(* IEC 61131-3 sources: iecf/harness/cases (part 3) *)

(* ---- locmore.st ---- *)
(* Located variables without a name (Ed.3 Loc_Var_Decl: Variable_Name ?)
   and a FOR control variable at an address. Worked by hand:
   AT %QW4 : INT := 5 sets %QW4 to 5 (Q bytes 4, 5: 05 00) as the
   program is set up; AT %MB0 : ARRAY [1..2] OF BYTE := [1, 2] sets
   %MB0, %MB1 (01 02); AT %QB9 : BYTE := 7 sets %QB9 (07) -
   in the PROGRAM: a block's VAR has no full address (Ed.3
   Other_Var_Decls).
   FOR i AT %MW2 := 1 TO 3 adds i to n: 6 (%QB0); i is 4 after it
   (%MW2, 04 00).
   FOR j AT %MW4 := 1 TO 5, left by EXIT at 3: j is 3 (%MW4, 03 00).
   FOR k AT %MW6 := 1 TO 10, the body adding 2 to k through a reference
   (assigned there itself it is E0015, Ed.3 7.3.3.4.2): k 1, 3; 4, 6; 7,
   9; 10, 12; then 13 is past 10: four passes (%QB1 4), k 13 (%MW6,
   0d 00).
   FOR z AT %MW8 := 5 TO 1 does not run: z is 5 (%MW8, 05 00).
   reference-skip: a located variable without a name, an array at an
   address: refused. *)
FUNCTION_BLOCK BT
  VAR n : INT; END_VAR
  n := n + 1;
END_FUNCTION_BLOCK
PROGRAM main
  VAR AT %QW4 : INT := 5; END_VAR
  VAR AT %MB0 : ARRAY [1..2] OF BYTE := [1, 2]; END_VAR
  VAR AT %QB9 : BYTE := 7; END_VAR
  VAR
    i AT %MW2 : INT;
    j AT %MW4 : INT;
    k AT %MW6 : INT;
    z AT %MW8 : INT;
    q0 AT %QB0 : SINT;
    q1 AT %QB1 : SINT;
  END_VAR
  VAR
    b : BT;
    n : INT;
    cnt : INT;
    rk : REF_TO INT;
  END_VAR
  b();
  n := 0;
  FOR i := 1 TO 3 DO
    n := n + i;
  END_FOR;
  q0 := INT_TO_SINT(n);
  FOR j := 1 TO 5 DO
    IF j = 3 THEN
      EXIT;
    END_IF;
  END_FOR;
  cnt := 0;
  rk := REF(k);
  FOR k := 1 TO 10 DO
    rk^ := rk^ + 2;
    cnt := cnt + 1;
  END_FOR;
  q1 := INT_TO_SINT(cnt);
  FOR z := 5 TO 1 DO
    cnt := 99;
  END_FOR;
END_PROGRAM

CONFIGURATION c
  RESOURCE r ON x
    TASK t(INTERVAL := T#10ms, PRIORITY := 1);
    PROGRAM p WITH t : main;
  END_RESOURCE
END_CONFIGURATION

(* ---- methods.st ---- *)
(* Methods and classes, bound statically (Ed.3 6.6.5, 6.6.7; OO.md step
   A): Ed.3's COUNTER (6.6.5.4.3 Example 2), UP5 calling THIS.UP; a
   method's result, its output taken, one without a result as a
   statement, one in an IF; a PUBLIC variable read and written from
   outside; a FUNCTION_BLOCK with a body and methods, the body calling
   THIS.Toggle, a method with in-outs; an input set from outside before
   the call; a method of an instance in an instance; EN on a method call.
   Worked amount hand, the input go at %IX0.0:
   tick 0, go FALSE: UP(3) CV 3 hits 1, q 3; UP5 CV 8 hits 2, q5 8, qf
   FALSE; not Full; qh 2, hits 12; L: lit FALSE (sw FALSE), then sw
   TRUE; Swap x 2 y 1, swaps.n 1, qx 21; Add(2) n 3, qs 3; EN FALSE: UP
   not called, qe stays 0.
   Tick 1, go TRUE: CV 11, 16, hits 13, 14; qh 14, hits 24; ql TRUE;
   qx 12, qs 6; UP(1) CV 17 hits 25, qe 17.
   Tick 2, go TRUE: UP(3) CV 20, q 20; UP5: 20 > 15, QU TRUE, q5 20, qf
   TRUE; Full: Reset, CV 0; hits 26, 27, qh 27, hits 37; qx 21, qs 9;
   UP(1) CV 1, qe 1.
   Tick 3, go FALSE: from CV 1, q 4, q5 9, qf FALSE, qh 40, ql FALSE, qx
   12, qs 12;
   qe stays 1.
   reference-skip: classes and methods are Ed.3's; the reference
   compiler (Ed.2) has neither. *)
CLASS COUNTER
  VAR CV : UINT; Top : UINT := 20; END_VAR
  VAR PUBLIC hits : INT; END_VAR
  METHOD PUBLIC UP : UINT
    VAR_INPUT INC : UINT; END_VAR
    VAR_OUTPUT QU : BOOL; END_VAR
    IF CV <= Top - INC THEN
      CV := CV + INC;
      QU := FALSE;
    ELSE
      QU := TRUE;
    END_IF;
    UP := CV;
    hits := hits + 1;
  END_METHOD
  METHOD PUBLIC UP5 : UINT
    VAR_OUTPUT QU : BOOL; END_VAR
    UP5 := THIS.UP(INC := 5, QU => QU);
  END_METHOD
  METHOD PUBLIC Full : BOOL
    Full := CV >= Top;
  END_METHOD
  METHOD PUBLIC Reset
    THIS.CV := 0;
  END_METHOD
END_CLASS

CLASS Tally
  VAR PUBLIC n : INT; END_VAR
  METHOD PUBLIC Add
    VAR_INPUT amount : INT := 1; END_VAR
    n := n + amount;
  END_METHOD
END_CLASS

FUNCTION_BLOCK Lamp
  VAR_INPUT sw : BOOL; END_VAR
  VAR_OUTPUT lit : BOOL; END_VAR
  VAR PUBLIC swaps : Tally; END_VAR
  METHOD PUBLIC Toggle
    sw := NOT sw;
  END_METHOD
  METHOD PUBLIC Swap
    VAR_IN_OUT a, b : INT; END_VAR
    VAR t : INT; END_VAR
    t := a;
    a := b;
    b := t;
    swaps.Add();
  END_METHOD
  lit := sw;
  THIS.Toggle();
END_FUNCTION_BLOCK

PROGRAM main
VAR
  CT : COUNTER;
  L : Lamp;
  lim : BOOL;
  x : INT := 1;
  y : INT := 2;
END_VAR
VAR
  go AT %IX0.0 : BOOL;
  q AT %QW0 : UINT;
  q5 AT %QW2 : UINT;
  qh AT %QW4 : INT;
  qx AT %QW6 : INT;
  qs AT %QW8 : INT;
  qf AT %QX10.0 : BOOL;
  ql AT %QX10.1 : BOOL;
  qe AT %QW11 : UINT;
END_VAR
q := CT.UP(INC := 3, QU => lim);
q5 := CT.UP5(QU => qf);
IF CT.Full() THEN
  CT.Reset();
END_IF;
qh := CT.hits;
CT.hits := CT.hits + 10;
L.sw := go;
L();
ql := L.lit;
L.Swap(a := x, b := y);
qx := x * 10 + y;
L.swaps.Add(amount := 2);
qs := L.swaps.n;
qe := CT.UP(EN := go, INC := 1);
END_PROGRAM

CONFIGURATION Plant
  RESOURCE r ON PLC
    TASK fast(INTERVAL := T#10ms, PRIORITY := 1);
    PROGRAM p WITH fast : main;
  END_RESOURCE
END_CONFIGURATION

(* ---- mutual.st ---- *)
(* Two blocks that name each other: b holds an a, and a takes a b as an
   in-out and through a reference, reads its output and calls its
   method. a's type is written before b's, which holds it; a's body
   after b's variables are known (docs/c-output.md §3). Worked by hand:

   tick 0: x(): total 0 + inner.n 0 + m 3 = 3 (Q2). y(other := x, r :=
   REF(x2)): n 0 + x.m 3 + x2.m 3 = 6 (Q0), and x2.poke(): 1 (Q4).
   tick 1: total 6; n 6 + 3 + 3 = 12 (0c 00); pokes 2.
   reference-skip: methods and REF_TO a block, as `refimage`. *)
FUNCTION_BLOCK a
  VAR_IN_OUT other : b; END_VAR
  VAR_INPUT r : REF_TO b; END_VAR
  VAR_OUTPUT n : INT; END_VAR
  n := n + other.m;
  IF r <> NULL THEN n := n + r^.m; r^.poke(); END_IF;
END_FUNCTION_BLOCK
FUNCTION_BLOCK b
  VAR inner : a; END_VAR
  VAR_OUTPUT m : INT := 3; total : INT; pokes : INT; END_VAR
  METHOD PUBLIC poke
    pokes := pokes + 1;
  END_METHOD
  total := total + inner.n + m;
END_FUNCTION_BLOCK
PROGRAM main
  VAR x : b; x2 : b; y : a; END_VAR
  VAR q AT %QW0 : ARRAY [0..2] OF INT; END_VAR
  x();
  y(other := x, r := REF(x2));
  q[0] := y.n;
  q[1] := x.total;
  q[2] := x2.pokes;
END_PROGRAM
CONFIGURATION c RESOURCE r ON PLC TASK t(INTERVAL := T#10ms, PRIORITY := 1); PROGRAM p WITH t : main; END_RESOURCE END_CONFIGURATION

(* ---- namespaces.st ---- *)
(* Namespaces (Ed.3 6.9; NAMESPACES.md), over two files: this one and
   namespaces.d/lib.st, which both add to the namespace Lib (Table 65
   NOTE).
   - Plant's own TON hides the standard one inside Plant (6.9.2
     Example 2): its ET is an INT that counts the calls with IN TRUE.
   - Plant's own area hides the one Plant's USING Lib.Shapes brings in
     (D2): w + h.
   - Lib.twice written inside Plant is Plant.Lib.twice, 3 x: the first
     part of a dotted name is found from inside out (D3).
   - outside, at global level, reaches Lib.Shapes.area through this
     file's USING (D6), area itself calls the INTERNAL offset of its own
     namespace, and Lib.tenfold calls Detail.scale, in the INTERNAL
     namespace Lib.Detail, from inside Lib (Figure 29).
   - Corner, a type of Lib.Shapes, by its short name through USING.
   Worked by hand, tick 0, vin 2: qa = area 2 + 3 = 5; qb = 3 * 2 = 6;
   qc = t.ET 1; qd = outside(2) = (2 * 2 + 100) + 2 * 2 + 2 * 10 = 128;
   qe = 7, c being Corner#Round.
   Tick 1, vin 5: qa 8; qb 15; qc 2; qd = (10 + 100) + 10 + 50 = 170;
   qe 7.
   reference-skip: the reference compiler (Ed.2) has no namespaces. *)
USING Lib.Shapes;

NAMESPACE Lib
    FUNCTION twice : INT
    VAR_INPUT x : INT; END_VAR
        twice := x * 2;
    END_FUNCTION
END_NAMESPACE

FUNCTION outside : INT
VAR_INPUT x : INT; END_VAR
    outside := area(x, 2) + Lib.twice(x) + Lib.tenfold(x);
END_FUNCTION

NAMESPACE Plant
    USING Lib.Shapes;

    FUNCTION_BLOCK TON
    VAR_INPUT IN : BOOL; END_VAR
    VAR_OUTPUT Q : BOOL; ET : INT; END_VAR
        IF IN THEN
            ET := ET + 1;
        END_IF;
        Q := ET >= 2;
    END_FUNCTION_BLOCK

    FUNCTION area : INT
    VAR_INPUT w, h : INT; END_VAR
        area := w + h;
    END_FUNCTION

    NAMESPACE Lib
        FUNCTION twice : INT
        VAR_INPUT x : INT; END_VAR
            twice := x * 3;
        END_FUNCTION
    END_NAMESPACE

    PROGRAM Main
    VAR
        vin AT %IW0 : INT;
        qa AT %QW0 : INT;
        qb AT %QW2 : INT;
        qc AT %QW4 : INT;
        qd AT %QW6 : INT;
        qe AT %QW8 : INT;
    END_VAR
    VAR
        t : TON;
        c : Corner := Corner#Round;
    END_VAR
        qa := area(vin, 3);
        qb := Lib.twice(vin);
        t(IN := TRUE);
        qc := t.ET;
        qd := outside(vin);
        IF c = Corner#Round THEN
            qe := 7;
        END_IF;
    END_PROGRAM
END_NAMESPACE

CONFIGURATION Works
  RESOURCE r ON PLC
    TASK fast(INTERVAL := T#10ms, PRIORITY := 1);
    PROGRAM p WITH fast : Plant.Main;
  END_RESOURCE
END_CONFIGURATION

(* ---- outelems.st ---- *)
(* Outputs of a structure, an array and a STRING type taken into an
   element by a computed index, and through a reference (Ed.3 6.6.1.4:
   Param_Assign, `Variable_Name '=>' Variable`): a FUNCTION's, found
   after it returns, and a function block's, found after it runs - the
   index checked there, as an elementary output's target is. Worked by
   hand: tick 0, i 1 (%IB0): Make(a := 5) into ps[1], ss[1], vs[1]:
   ps[1].x 5 (%QB0), ps[1].y 10 (%QB1), vs[1][1] 7 (%QB2), ss[1] 'ab'
   (%QX7.0); g(a := 7) into ps[2], ss[2]: ps[2].x 7 (%QB3), ps[2].y -7
   (%QB4), ss[2] 'cd' (%QX7.1); Make(a := 3) through rp^ and rst^ into pnt
   and st: pnt.x 3 (%QB5), pnt.y 6 (%QB6), st 'ab' (%QX7.2). Last, a
   whole output of an instance that is an element read, pnt :=
   gs[i - 1].p after gs[0](a := 4): 4 (%QB8), -4 (%QB9).
   Tick 1, i 2: Make into ps[2] (5, 10), then g's target ps[3] is
   outside 0..2: the task stops there, fault INDEX, line 70, after g
   ran and before its outputs are stored.
   reference-skip: the reference compiler refuses REF_TO STRING[8], and
   its C for an output into an element does not compile (as fnoutx). *)
TYPE POINT : STRUCT x, y : INT; END_STRUCT; END_TYPE

FUNCTION Make : INT
  VAR_INPUT a : INT; END_VAR
  VAR_OUTPUT p : POINT; s : STRING[8]; v : ARRAY[0..1] OF INT; END_VAR
  p.x := a;
  p.y := a * 2;
  s := 'ab';
  v[0] := a + 1;
  v[1] := a + 2;
  Make := a;
END_FUNCTION

FUNCTION_BLOCK Gen
  VAR_INPUT a : INT; END_VAR
  VAR_OUTPUT p : POINT; s : STRING[8]; END_VAR
  p.x := a;
  p.y := -a;
  s := 'cd';
END_FUNCTION_BLOCK

PROGRAM main
  VAR
    i AT %IB0 : SINT;
  END_VAR
  VAR
    ps : ARRAY[0..2] OF POINT;
    ss : ARRAY[0..2] OF STRING[8];
    vs : ARRAY[0..2] OF ARRAY[0..1] OF INT;
    g : Gen;
    gs : ARRAY[0..1] OF Gen;
    pnt : POINT;
    st : STRING[8];
    rp : REF_TO POINT;
    rst : REF_TO STRING[8];
    n : INT;
  END_VAR
  VAR
    q0 AT %QB0 : SINT;
    q1 AT %QB1 : SINT;
    q2 AT %QB2 : SINT;
    q3 AT %QB3 : SINT;
    q4 AT %QB4 : SINT;
    q5 AT %QB5 : SINT;
    q6 AT %QB6 : SINT;
    c0 AT %QX7.0 : BOOL;
    c1 AT %QX7.1 : BOOL;
    c2 AT %QX7.2 : BOOL;
    q8 AT %QB8 : SINT;
    q9 AT %QB9 : SINT;
  END_VAR
  n := Make(a := 5, p => ps[i], s => ss[i], v => vs[i]);
  g(a := 7, p => ps[i + 1], s => ss[i + 1]);
  rp := REF(pnt);
  rst := REF(st);
  n := Make(a := 3, p => rp^, s => rst^);
  q0 := INT_TO_SINT(ps[1].x);
  q1 := INT_TO_SINT(ps[1].y);
  q2 := INT_TO_SINT(vs[1][1]);
  q3 := INT_TO_SINT(ps[2].x);
  q4 := INT_TO_SINT(ps[2].y);
  q5 := INT_TO_SINT(pnt.x);
  q6 := INT_TO_SINT(pnt.y);
  c0 := ss[1] = 'ab';
  c1 := ss[2] = 'cd';
  c2 := st = 'ab';
  gs[i - 1](a := 4);
  pnt := gs[i - 1].p;
  q8 := INT_TO_SINT(pnt.x);
  q9 := INT_TO_SINT(pnt.y);
END_PROGRAM

CONFIGURATION c
  RESOURCE r ON x
    TASK t(INTERVAL := T#10ms, PRIORITY := 1);
    PROGRAM p WITH t : main;
  END_RESOURCE
END_CONFIGURATION

(* ---- partaccess.st ---- *)
(* Partial access of bit strings (Ed.3 6.6.1.3, Table 17): a bit, byte,
   word or double word of a BYTE, WORD, DWORD or LWORD, numbered from
   the least significant; read, and written into its whole. Worked by
   hand:
   w 16#1234: w.2 is TRUE (%QX0.0). w.%X0 := TRUE makes 16#1235;
   w.%B1 is 16#12 (%QB1). w.%B0 := 16#FF makes 16#12FF: %QB2 FF, %QB3
   12.
   dw 16#AABBCCDD: w2 := dw.%W1 is 16#AABB: %QB4 BB, %QB5 AA.
   dw.%W0 := 16#1122 makes 16#AABB1122: dw.%B0 22 (%QB6).
   l 0: l.63 := TRUE, l.%D0 := 16#01020304: l.%B7 80 (%QB7), l.%B2 02
   (%QB8).
   a[i].3 := TRUE with i 2: a[2] 8 (%QB9).
   m AT %MW0: m.%B1 := 16#AB writes its high byte, %MB1 (the M bytes
   00 AB); m.15 is TRUE (%QX10.0).
   r := REF(w); r^.%B1 := 16#77: w 16#77FF, w.%B1 77 (%QB11).
   o(q => w.0), q FALSE: w 16#77FE, w.%B0 FE (%QB12).
   Last, a[i].0 := TRUE with i 3: the index faults (INDEX) before the
   store.
   reference-skip: the reference compiler (Ed.2) has no partial
   access. *)
FUNCTION_BLOCK OT
  VAR_OUTPUT q : BOOL; END_VAR
  q := FALSE;
END_FUNCTION_BLOCK
PROGRAM main
  VAR
    w : WORD := 16#1234;
    w2 : WORD;
    dw : DWORD := 16#AABBCCDD;
    l : LWORD;
    a : ARRAY [1..2] OF WORD;
    i : INT := 2;
    r : REF_TO WORD;
    o : OT;
  END_VAR
  VAR
    m AT %MW0 : WORD;
    q00 AT %QX0.0 : BOOL;
    q1 AT %QB1 : BYTE;
    q2 AT %QB2 : BYTE;
    q3 AT %QB3 : BYTE;
    q4 AT %QB4 : BYTE;
    q5 AT %QB5 : BYTE;
    q6 AT %QB6 : BYTE;
    q7 AT %QB7 : BYTE;
    q8 AT %QB8 : BYTE;
    q9 AT %QB9 : BYTE;
    q10 AT %QX10.0 : BOOL;
    q11 AT %QB11 : BYTE;
    q12 AT %QB12 : BYTE;
  END_VAR
  q00 := w.2;
  w.%X0 := TRUE;
  q1 := w.%B1;
  w.%B0 := 16#FF;
  q2 := w.%B0;
  q3 := w.%B1;
  w2 := dw.%W1;
  q4 := w2.%B0;
  q5 := w2.%B1;
  dw.%W0 := 16#1122;
  q6 := dw.%B0;
  l.63 := TRUE;
  l.%D0 := 16#01020304;
  q7 := l.%B7;
  q8 := l.%B2;
  a[i].3 := TRUE;
  q9 := a[2].%B0;
  m.%B1 := 16#AB;
  q10 := m.15;
  r := REF(w);
  r^.%B1 := 16#77;
  q11 := w.%B1;
  o(q => w.0);
  q12 := w.%B0;
  i := 3;
  a[i].0 := TRUE;
END_PROGRAM

CONFIGURATION c
  RESOURCE r ON x
    TASK t(INTERVAL := T#10ms, PRIORITY := 1);
    PROGRAM p WITH t : main;
  END_RESOURCE
END_CONFIGURATION

(* ---- partlyoutput.st ---- *)
(* A function block's VAR_OUTPUT of a structure with `*` components
   (Ed.3 6.4.4.8 excludes only VAR_INPUT, VAR_IN_OUT and VAR_TEMP),
   completed per instance by VAR_CONFIG (6.5.5.4): d.o.q at %QW0, d.o.m
   at %MW0; the program's own s of the same type at %QW2 and %MW2.
   Worked by hand, k counting 1, 2: d sets o.q := n * 2, o.m + 1; the
   program reads d.o.m into %QW4 and copies d.o into s.
   Tick 0: %QW0 2, %QW2 2, %QW4 1; %MW0 1, %MW2 1.
   Tick 1: %QW0 4, %QW2 4, %QW4 2; %MW0 2, %MW2 2.
   reference-skip: the reference compiler has no `*` structure components. *)
TYPE Out : STRUCT
  q AT %Q* : INT;
  m AT %M* : INT;
END_STRUCT;
END_TYPE

FUNCTION_BLOCK Drive
  VAR_INPUT n : INT; END_VAR
  VAR_OUTPUT o : Out; END_VAR
  o.q := n * 2;
  o.m := o.m + 1;
END_FUNCTION_BLOCK

PROGRAM main
  VAR d : Drive; k : INT; s : Out; END_VAR
  VAR seen AT %QW4 : INT; END_VAR
  k := k + 1;
  d(n := k);
  seen := d.o.m;
  s := d.o;
END_PROGRAM

CONFIGURATION cf
  RESOURCE rs ON x
    TASK tk(INTERVAL := T#10ms, PRIORITY := 1);
    PROGRAM p WITH tk : main;
  END_RESOURCE
  VAR_CONFIG
    rs.p.d.o.q AT %QW0 : INT;
    rs.p.d.o.m AT %MW0 : INT;
    rs.p.s.q AT %QW2 : INT;
    rs.p.s.m AT %MW2 : INT;
  END_VAR
END_CONFIGURATION

(* ---- pous.st ---- *)
(* The user's POUs: a FUNCTION with inputs by name and by position, a
   FUNCTION_BLOCK keeping state across ticks, VAR_IN_OUT, VAR_OUTPUT read
   from outside, an FB instance inside an FB, and globals of the
   CONFIGURATION through VAR_EXTERNAL. *)
FUNCTION scale : INT
VAR_INPUT
  x : INT;
  num : INT := 1;
  den : INT := 1;
END_VAR
scale := x * num / den;
END_FUNCTION

FUNCTION_BLOCK average
VAR_INPUT
  sample : INT;
END_VAR
VAR_OUTPUT
  avg : INT;
  count : INT;
END_VAR
VAR
  sum : DINT;
END_VAR
sum := sum + INT_TO_DINT(sample);
count := count + 1;
avg := DINT_TO_INT(sum / INT_TO_DINT(count));
END_FUNCTION_BLOCK

FUNCTION_BLOCK twice
VAR_IN_OUT
  v : INT;
END_VAR
VAR_OUTPUT
  inner_avg : INT;
END_VAR
VAR
  a : average;
END_VAR
v := v * 2;
a(sample := v);
inner_avg := a.avg;
END_FUNCTION_BLOCK

PROGRAM main
VAR
  inp AT %IW0 : INT;
  r_pos AT %MW0 : INT;
  r_named AT %MW2 : INT;
  r_default AT %MW4 : INT;
  r_avg AT %MW6 : INT;
  r_count AT %MW8 : INT;
  r_inout AT %MW10 : INT;
  r_inner AT %MW12 : INT;
  r_global AT %MW14 : INT;
END_VAR
VAR
  avg1 : average;
  tw : twice;
  local : INT := 1;
END_VAR
VAR_EXTERNAL
  g_total : INT;
END_VAR
VAR_EXTERNAL CONSTANT
  g_limit : INT;
END_VAR
r_pos := scale(inp, 3, 2);
r_named := scale(den := 4, x := inp, num := 2);
r_default := scale(x := inp);
avg1(sample := inp);
r_avg := avg1.avg;
r_count := avg1.count;
tw(v := local);
r_inout := local;
r_inner := tw.inner_avg;
IF g_total < g_limit THEN
  g_total := g_total + inp;
END_IF;
r_global := g_total;
END_PROGRAM

CONFIGURATION plant
  VAR_GLOBAL
    g_total : INT := 0;
  END_VAR
  VAR_GLOBAL CONSTANT
    g_limit : INT := 50;
  END_VAR
  RESOURCE r ON PLC
    TASK fast(INTERVAL := T#10ms, PRIORITY := 0);
    PROGRAM p WITH fast : main;
  END_RESOURCE
END_CONFIGURATION

(* ---- prginst.st ---- *)
(* Programs as single instances (the program-instances extension), as
   CODESYS and TwinCAT have them. counter runs in its task with inc 1
   and total to sum, and main, after it, calls it with inc 100, calls
   its method Bump(1) and adds 10 to its calls: one instance, shared.
   Worked by hand: tick 0 - the task: total 1, calls 1, sum 1; main:
   total 101, calls 2, Bump 102, calls 12. Tick 1: total 103, calls 13,
   sum 103; 203, 14, 204, 24. Tick 2: 205, 25, 205; 305, 26, 306, 36.
   So %QB1 (calls) 12 24 36, %QB2 (Bump MOD 100) 2 4 6, %QB3 (sum MOD
   100) 1 3 5. NO.v is NO's v, not a value of E1 or E2: h's FB_init
   took it, 6, as h was set up (%QB0); main adds 1 each tick, %QB4 7 8
   9; e keeps E2#No (%QB5 1).
   reference-skip: a program read and called by its name is CODESYS's,
   not IEC 61131-3. *)
{attribute 'qualified_only'}
TYPE E1 : (No := 1, Yes := 2); END_TYPE
{attribute 'qualified_only'}
TYPE E2 : (No := 3, Maybe := 4); END_TYPE

PROGRAM NO
VAR v : INT := 6; END_VAR
END_PROGRAM

PROGRAM counter
VAR_INPUT inc : INT; END_VAR
VAR_OUTPUT total : INT; END_VAR
VAR calls : INT; END_VAR
METHOD Bump : INT
VAR_INPUT n : INT; END_VAR
total := total + n;
Bump := total;
END_METHOD
total := total + inc;
calls := calls + 1;
END_PROGRAM

FUNCTION_BLOCK Holder
VAR_OUTPUT got : INT; END_VAR
METHOD FB_init : BOOL
VAR_INPUT bInitRetains : BOOL; bInCopyCode : BOOL; start : INT; END_VAR
got := start;
END_METHOD
END_FUNCTION_BLOCK

PROGRAM main
VAR h : Holder(NO.v); r : INT; e : E2 := E2.No; END_VAR
VAR_EXTERNAL sum : INT; END_VAR
VAR q0 AT %QB0 : SINT; q1 AT %QB1 : SINT; q2 AT %QB2 : SINT; q3 AT %QB3 : SINT; q4 AT %QB4 : SINT;
    q5 AT %QB5 : SINT; END_VAR
counter(inc := 100);
r := counter.Bump(1);
counter.calls := counter.calls + 10;
NO.v := NO.v + 1;
q0 := INT_TO_SINT(h.got);
q1 := INT_TO_SINT(counter.calls);
q2 := INT_TO_SINT(r MOD 100);
q3 := INT_TO_SINT(sum MOD 100);
q4 := INT_TO_SINT(NO.v);
q5 := BOOL_TO_SINT(e = E2.No);
END_PROGRAM

CONFIGURATION cf
  VAR_GLOBAL sum : INT; END_VAR
  RESOURCE r ON x
    TASK tk(INTERVAL := T#10ms, PRIORITY := 1);
    PROGRAM c WITH tk : counter(inc := 1, total => sum);
    PROGRAM m WITH tk : main;
  END_RESOURCE
END_CONFIGURATION

(* ---- progglobals.st ---- *)
(* A PROGRAM's own VAR_GLOBAL (Ed.3 Table 47, 8a and 8b): each instance
   of the program has its own, seen by the instances it holds and the
   FUNCTIONs it calls. main runs twice in r1, a and b, each with its own
   z, gi and kept; solo has a z of its own, which its FUNCTION reads;
   plain, in r2, reaches r2's z. Worked by hand, inc 2:

   tick 0, a (z 5): c 7, the VAR_TEMP t 9, h.c 11, gi, the program's
   global instance, 13, v's own VAR_TEMP 15; z + 10 = 25 (Q0 19 00); q2
   13 + 15 = 28 (Q2 1c 00); kept 51 (Q4 33). b: the same, of its own
   (Q8 19 00, Q10 1c 00, Q12 33). out is at %QB20 for both: 2. solo (z
   1000, then VAR_CONFIG's 2000): c 2002, readz 2002 (Q16 d2 07). plain (r2's z 300): 302 (Q18
   2e 01).
   tick 1, a (z 25): 27, 29, 31, 33, 35; 45 (2d 00); 33 + 35 = 68 (44
   00); kept 52. solo 2004, plain 304, out 4.
   warm, before tick 2: all starts again but kept, RETAIN, each
   instance's own (53), and out, in the image (6).
   reference-skip: VAR_GLOBAL in a PROGRAM: the reference compiler
   refuses it. *)
TYPE Hold : STRUCT c : counter; END_STRUCT; END_TYPE
FUNCTION_BLOCK counter
  VAR_EXTERNAL z : INT; END_VAR
  VAR_EXTERNAL CONSTANT inc : INT; END_VAR
  VAR_OUTPUT o : INT; END_VAR
  z := z + inc;
  o := z;
END_FUNCTION_BLOCK
FUNCTION readz : INT
  VAR_EXTERNAL z : INT; END_VAR
  readz := z;
END_FUNCTION
FUNCTION_BLOCK viatemp
  VAR_OUTPUT o : INT; END_VAR
  VAR_TEMP t : counter; END_VAR
  t();
  o := t.o;
END_FUNCTION_BLOCK
PROGRAM main
  VAR_GLOBAL z : INT := 5; gi : counter; END_VAR
  VAR_GLOBAL CONSTANT inc : INT := 2; END_VAR
  VAR_GLOBAL RETAIN kept : USINT := 50; END_VAR
  VAR_GLOBAL out AT %QB20 : USINT; END_VAR
  VAR c : counter; h : Hold; v : viatemp; END_VAR
  VAR q AT %Q* : INT; q2 AT %Q* : INT; q3 AT %Q* : USINT; END_VAR
  VAR_TEMP t : counter; END_VAR
  c();
  t();
  h.c();
  gi();
  v();
  z := z + 10;
  q := z;
  q2 := gi.o + v.o;
  kept := kept + 1;
  q3 := kept;
  out := out + 1;
END_PROGRAM
PROGRAM solo
  VAR_GLOBAL z : INT := 1000; END_VAR
  VAR_GLOBAL CONSTANT inc : INT := 2; END_VAR
  VAR c : counter; END_VAR
  VAR q AT %QW16 : INT; END_VAR
  c();
  q := readz();
END_PROGRAM
PROGRAM plain
  VAR c : counter; END_VAR
  VAR q AT %QW18 : INT; END_VAR
  c();
  q := c.o;
END_PROGRAM
CONFIGURATION plant
  RESOURCE r1 ON PLC
    TASK t(INTERVAL := T#10ms, PRIORITY := 1);
    PROGRAM a WITH t : main;
    PROGRAM b WITH t : main;
    PROGRAM s WITH t : solo;
  END_RESOURCE
  RESOURCE r2 ON PLC
    VAR_GLOBAL z : INT := 300; END_VAR
    VAR_GLOBAL CONSTANT inc : INT := 2; END_VAR
    TASK t(INTERVAL := T#10ms, PRIORITY := 2);
    PROGRAM p WITH t : plain;
  END_RESOURCE
  VAR_CONFIG
    r1.a.q AT %QW0 : INT;
    r1.a.q2 AT %QW2 : INT;
    r1.a.q3 AT %QB4 : USINT;
    r1.b.q AT %QW8 : INT;
    r1.b.q2 AT %QW10 : INT;
    r1.b.q3 AT %QB12 : USINT;
    r1.s.z : INT := 2000;
  END_VAR
END_CONFIGURATION

(* ---- progretain.st ---- *)
(* RETAIN on a program instance (Ed.3 6.5.6.2): the instance's variables
   of sections neither RETAIN nor NON_RETAIN are kept across a warm
   restart; one that is itself a block keeps what its own type says. a
   is RETAIN, b is plain, c NON_RETAIN, which is what b is. o is a + p.x
   + arr[1] + c.n + c.kept + r + nr + LEN(s). Worked by hand:

   init: ini 7 at each instance's address, VAR_CONFIG's (Q2, Q6, Q10).
   tick 0, a (VAR_CONFIG's a 100, inc 1): 101 + 4 + 7 + 1 + 1 + 21 + 31
   + 3 = 169 (Q0 a9 00, and oa, Q20); ini 8. b (a 200, inc 2): 202 + 4 +
   7 + 1 + 1 + 21 + 31 + 3 = 270 (Q4 0e 01, ob, Q22). c (a 10): 11 + ...
   = 79 (Q8 4f 00).
   tick 1: a 102 + 5 + 8 + 2 + 2 + 22 + 32 + 4 = 177 (b1 00), ini 9; b
   204 + ... = 279 (17 01); c 87 (57 00).
   warm, before tick 2. a keeps a 102 (VAR_CONFIG's 100 is not given
   again), p.x 5, arr[1] 8, s 'abxx', inc, and ini, 9, in the image; r is
   RETAIN anyway; nr, NON_RETAIN, starts at 30; its block c starts again
   but for its own RETAIN kept, 2. b and c keep r and the block's kept
   alone: a 200 and 10 again, ini 7.
   tick 2: a 103 + 6 + 9 + 1 + 3 + 23 + 31 + 5 = 181 (b5 00), ini 10; b
   202 + 4 + 7 + 1 + 3 + 23 + 31 + 3 = 274 (12 01), ini 8; c 83 (53 00).
   tick 3: a 104 + 7 + 10 + 2 + 4 + 24 + 32 + 6 = 189 (bd 00), ini 11; b
   283 (1b 01); c 91 (5b 00).
   reference-skip: AT %Q* in a PROGRAM; VAR_CONFIG generates nothing;
   no warm restart. *)
TYPE Pt : STRUCT x : INT := 3; y : INT; END_STRUCT; END_TYPE
FUNCTION_BLOCK counter
  VAR_OUTPUT n : INT; END_VAR
  VAR_OUTPUT RETAIN kept : INT; END_VAR
  n := n + 1;
  kept := kept + 1;
END_FUNCTION_BLOCK
PROGRAM main
  VAR_INPUT inc : INT := 1; END_VAR
  VAR a : INT := 10; p : Pt; arr : ARRAY [0..1] OF INT := [5, 6]; c : counter; tm : TON; s : STRING[8] := 'ab'; END_VAR
  VAR RETAIN r : INT := 20; END_VAR
  VAR NON_RETAIN nr : INT := 30; END_VAR
  VAR q AT %Q* : INT; END_VAR
  VAR ini AT %Q* : INT; END_VAR
  VAR_OUTPUT o : INT; END_VAR
  a := a + inc;
  p.x := p.x + 1;
  arr[1] := arr[1] + 1;
  c();
  r := r + 1;
  nr := nr + 1;
  ini := ini + 1;
  s := CONCAT(s, 'x');
  o := a + p.x + arr[1] + c.n + c.kept + r + nr + LEN(s);
  q := o;
END_PROGRAM
CONFIGURATION plant
  VAR_GLOBAL two : INT := 2; oa AT %QW20 : INT; ob AT %QW22 : INT; END_VAR
  RESOURCE cpu ON PLC
    TASK t(INTERVAL := T#10ms, PRIORITY := 1);
    PROGRAM RETAIN a WITH t : main(o => oa);
    PROGRAM b WITH t : main(inc := two, o => ob);
    PROGRAM NON_RETAIN c WITH t : main;
  END_RESOURCE
  VAR_CONFIG
    cpu.a.q AT %QW0 : INT;
    cpu.a.ini AT %QW2 : INT := 7;
    cpu.b.q AT %QW4 : INT;
    cpu.b.ini AT %QW6 : INT := 7;
    cpu.c.q AT %QW8 : INT;
    cpu.c.ini AT %QW10 : INT := 7;
    cpu.a.a : INT := 100;
    cpu.b.a : INT := 200;
  END_VAR
END_CONFIGURATION

(* ---- querypointer.st ---- *)
(* __QUERYPOINTER (the query-pointer extension): the instance an
   interface refers to as a POINTER TO its block - a reference to it -
   its type checked, where CODESYS leaves it to the program. Worked by
   hand: i a Lamp, w 3: TRUE, p^.w 3 (%QB0 1, %QB1 3); a BigLamp, derived
   from Lamp, w 5: TRUE, 5 (%QB2 5); a Motor, another type: FALSE and p
   0 (%QB3 10); NULL: FALSE (%QB4 0); q := ADR(l), q^.w := 9 writes l's w
   (%QB5 9); then p, 0, read: IECF_FAULT_NULL on line 50, %QB6 left 1.
   reference-skip: __QUERYPOINTER is CODESYS's, not IEC 61131-3. *)
INTERFACE IShape
METHOD Area : INT
END_METHOD
END_INTERFACE

FUNCTION_BLOCK Lamp IMPLEMENTS IShape
VAR_INPUT w : INT; END_VAR
METHOD PUBLIC Area : INT
Area := w;
END_METHOD
END_FUNCTION_BLOCK

FUNCTION_BLOCK BigLamp EXTENDS Lamp
END_FUNCTION_BLOCK

FUNCTION_BLOCK Motor IMPLEMENTS IShape
VAR_INPUT r : INT; END_VAR
METHOD PUBLIC Area : INT
Area := r;
END_METHOD
END_FUNCTION_BLOCK

PROGRAM main
VAR l : Lamp := (w := 3); b : BigLamp := (w := 5); m : Motor := (r := 7); i : IShape;
    p, q : POINTER TO Lamp; ok : BOOL; END_VAR
VAR q0 AT %QB0 : SINT; q1 AT %QB1 : SINT; q2 AT %QB2 : SINT; q3 AT %QB3 : SINT; q4 AT %QB4 : SINT;
    q5 AT %QB5 : SINT; q6 AT %QB6 : SINT; END_VAR
i := l;
q0 := BOOL_TO_SINT(__QUERYPOINTER(i, p));
q1 := INT_TO_SINT(p^.w);
i := b;
IF __QUERYPOINTER(i, p) THEN q2 := INT_TO_SINT(p^.w); END_IF;
i := m;
ok := __QUERYPOINTER(i, p);
q3 := BOOL_TO_SINT(ok) + 10 * BOOL_TO_SINT(p = 0);
i := NULL;
q4 := BOOL_TO_SINT(__QUERYPOINTER(i, p));
q := ADR(l);
q^.w := 9;
q5 := INT_TO_SINT(l.w);
q6 := 1;
q6 := INT_TO_SINT(p^.w);
END_PROGRAM

CONFIGURATION cf
  RESOURCE r ON x
    TASK tk(INTERVAL := T#10ms, PRIORITY := 1);
    PROGRAM pm WITH tk : main;
  END_RESOURCE
END_CONFIGURATION

(* ---- recursion.st ---- *)
(* A FUNCTION, a method and a block's body calling themselves
   (recursion), each call counted. Worked by hand:
   %QD0: fact(10), 3628800 (16#375F00), 00 5f 37 00.
   %QW4: t's o, sum(4) = 4 + 3 + 2 + 1, 10, 0a 00.
   %QW6: c's o, one for each of its three calls of itself, 03 00.
   %QD8: runaway(0) calls itself without an end: the call past
   IECF_DEPTH_MAX (64) is a fault, 14 (IECF_FAULT_DEPTH), at runaway's
   line 19, and %QD8 stays 0.
   reference-skip: the reference compiler knows a POU only after its
   declaration, so it can express no recursion. *)
FUNCTION fact : DINT
  VAR_INPUT n : DINT; END_VAR
  IF n <= 1 THEN fact := 1; RETURN; END_IF;
  fact := n * fact(n - 1);
END_FUNCTION

FUNCTION runaway : DINT
  VAR_INPUT n : DINT; END_VAR
  runaway := runaway(n + 1);
END_FUNCTION

FUNCTION_BLOCK Tree
  VAR_INPUT n : INT; END_VAR
  VAR_OUTPUT o : INT; END_VAR
  METHOD sum : INT
    VAR_INPUT k : INT; END_VAR
    IF k = 0 THEN sum := 0; RETURN; END_IF;
    sum := k + THIS.sum(k - 1);
  END_METHOD
  o := THIS.sum(n);
END_FUNCTION_BLOCK

FUNCTION_BLOCK Count
  VAR_INPUT n : INT; END_VAR
  VAR_IN_OUT me : Count; END_VAR
  VAR_OUTPUT o : INT; END_VAR
  IF n > 0 THEN
    o := o + 1;
    me(n := n - 1, me := me);
  END_IF;
END_FUNCTION_BLOCK

PROGRAM main
  VAR t : Tree; c : Count; END_VAR
  VAR q AT %QD0 : DINT; w AT %QW4 : INT; v AT %QW6 : INT; r AT %QD8 : DINT; END_VAR
  q := fact(10);
  t(n := 4);
  w := t.o;
  c(n := 3, me := c);
  v := c.o;
  r := runaway(0);
END_PROGRAM

CONFIGURATION cf
  RESOURCE r ON x
    TASK tk(INTERVAL := T#10ms, PRIORITY := 1);
    PROGRAM p WITH tk : main;
  END_RESOURCE
END_CONFIGURATION

(* ---- refimage.st ---- *)
(* References into the process image, to function blocks, and to
   references (Ed.3 6.4.4.10; docs/c-output.md §4): REF() of a variable
   at an address - a word, a BOOL at a bit, a BOOL taking a whole byte,
   an array, a structure, a STRING, an input - read and written through
   `^` as the variable itself is; REF() as an initial value; `r^ := ...`;
   an array of references and a reference to one, `rr^^`; a block, the
   user's and a standard one, called and read through a reference; a
   structure referencing its own type; `=` with REF(). At tick 5 %IW0 is
   99 and a NULL reference is dereferenced: a fault (IECF_FAULT_NULL), the
   statement stores nothing, and the task stops, as at tick 6.
   reference-skip: the reference compiler's C for `r^ := ...` does not
   compile, REF_TO a function block crashes it, and it has no REF() in an
   initial value or a comparison. *)
TYPE
  pair : STRUCT a : INT; b : BYTE; END_STRUCT;
  rint : REF_TO INT;
  node : STRUCT v : INT; next : REF_TO node; END_STRUCT;
END_TYPE

FUNCTION_BLOCK acc
VAR_INPUT x : INT; END_VAR
VAR_OUTPUT total : INT; END_VAR
total := total + x;
END_FUNCTION_BLOCK

PROGRAM main
VAR
  vin AT %IW0 : INT;
END_VAR
VAR
  w AT %MW0 : INT;
  bx AT %MX2.3 : BOOL;
  bb AT %MB3 : BOOL;
  la AT %MW4 : ARRAY[0..2] OF INT;
  ls AT %MW10 : pair;
  s AT %MB13 : STRING[3];
  o_tot AT %MW17 : INT;
  o_cnt AT %MW19 : INT;
  o_q AT %MX21.0 : BOOL;
  o_eq AT %MX21.1 : BOOL;
  o_node AT %MW22 : INT;
  o_pick AT %MW24 : INT;
  o_kept AT %MW26 : INT;
END_VAR
VAR
  rw : rint := REF(w);
  rin : REF_TO INT := REF(vin);
  rbx, rbb : REF_TO BOOL;
  rla : REF_TO ARRAY[0..2] OF INT;
  rls : REF_TO pair;
  rstr : REF_TO STRING[3];
  refs : ARRAY[0..2] OF rint;
  rr : REF_TO rint;
  k, kept : INT;
  f : acc;
  rf : REF_TO acc;
  c : CTU;
  rc : REF_TO CTU;
  n1, n2 : node;
  rn : REF_TO node;
END_VAR
k := vin MOD 3;
IF k < 0 THEN
  k := k + 3;
END_IF;
rw^ := rw^ + rin^;
rbx := REF(bx);
rbx^ := NOT rbx^;
rbb := REF(bb);
rbb^ := vin > 1;
rla := REF(la);
rla^[k] := rla^[k] + 10;
rls := REF(ls);
rls^.a := w;
rls^.b := INT_TO_BYTE(k);
rstr := REF(s);
IF k = 0 THEN
  rstr^ := 'ab';
ELSIF k = 1 THEN
  rstr^ := 'xyz';
ELSE
  rstr^ := '';
END_IF;
refs[0] := REF(la[0]);
refs[1] := REF(la[1]);
refs[2] := REF(la[2]);
rr := REF(refs[k]);
o_pick := rr^^;
rf := REF(f);
rf^(x := k + 1);
o_tot := rf^.total;
rc := REF(c);
rc^(CU := NOT rc^.CU, PV := 3);
o_cnt := rc^.CV;
o_q := rc^.Q;
o_eq := rw = REF(w);
n1.next := REF(n2);
n1.next^.v := n1.next^.v + k;
o_node := n2.v;
IF vin = 99 THEN
  rn := NULL;
ELSE
  rn := REF(n1);
END_IF;
kept := kept + 1;
o_kept := kept;
o_kept := rn^.v;
END_PROGRAM

CONFIGURATION c
  RESOURCE r ON PLC
    TASK t(INTERVAL := T#10ms, PRIORITY := 1);
    PROGRAM inst WITH t : main;
  END_RESOURCE
END_CONFIGURATION

(* ---- refmore.st ---- *)
(* References a FUNCTION gives (Ed.3 6.4.4.10), stored through and
   called through; a block's input and a whole instance set through a
   reference; a standard block's input set from outside (Ed.3 6.6.7.2.2,
   Figure 20 a); REF() of an interface variable.
   g1 1, g2 2. Pick(w) gives REF(g2) if w, else REF(g1). Worked by hand:
   r := Pick(TRUE): r^ 2 (%QB0). Pick(FALSE)^ := 5 writes g1: 5 (%QB1).
   Nul() sets no result: NULL (%QB2 1).
   PickP()^.x := 7 writes gp.x: 7 (%QB3); PickP()^.x + 1: 8 (%QB4).
   PickB()^.i := 3; PickB()^() adds i to n: gb.n 3 (%QB5).
   PickB()^(i := 4); PickB()^.n: 7 (%QB6).
   rb := REF(gb); rb^ := b2, a copy of b2, whose i is 10 and n 0; then
   gb() adds 10: gb.n 10 (%QB7).
   tm.PT := T#2s, set from outside: T#2s (%QB8 1). rt := REF(gt1);
   rt^.PT := T#3s: gt1.PT T#3s (%QB9 1). PickT()^.PT := T#4s: T#4s
   (%QB10 1). t3.PT := T#9s; rt^ := t3 copies t3 into gt1: T#9s (%QB11
   1).
   o1 gives 3, o2 6. pi := REF(i); pi^ := o1: i.g() 3 (%QB12).
   pi := REF(is[2]); pi^ := o2: is[2].g() 6 (%QB13), and pi^ is not
   NULL (%QB14 1).
   Last, Nul()^ read: NULL dereferenced faults NULL, nothing stored
   (%QB15 stays 0).
   reference-skip: methods; a write through a reference: its C does
   not build. *)
TYPE
  PT : STRUCT x : INT; END_STRUCT;
END_TYPE
INTERFACE IG
  METHOD g : INT END_METHOD
END_INTERFACE
FUNCTION_BLOCK BG IMPLEMENTS IG
  VAR_INPUT n : INT; END_VAR
  METHOD PUBLIC g : INT
    g := n;
  END_METHOD
END_FUNCTION_BLOCK
FUNCTION_BLOCK BA
  VAR_INPUT i : INT; END_VAR
  VAR_OUTPUT n : INT; END_VAR
  n := n + i;
END_FUNCTION_BLOCK
FUNCTION Pick : REF_TO INT
  VAR_INPUT w : BOOL; END_VAR
  VAR_EXTERNAL g1 : INT; g2 : INT; END_VAR
  IF w THEN
    Pick := REF(g2);
  ELSE
    Pick := REF(g1);
  END_IF;
END_FUNCTION
FUNCTION PickP : REF_TO PT
  VAR_EXTERNAL gp : PT; END_VAR
  PickP := REF(gp);
END_FUNCTION
FUNCTION PickB : REF_TO BA
  VAR_EXTERNAL gb : BA; END_VAR
  PickB := REF(gb);
END_FUNCTION
FUNCTION PickT : REF_TO TON
  VAR_EXTERNAL gt1 : TON; END_VAR
  PickT := REF(gt1);
END_FUNCTION
FUNCTION Nul : REF_TO INT
END_FUNCTION
PROGRAM main
  VAR_EXTERNAL g1 : INT; g2 : INT; gp : PT; gb : BA; gt1 : TON; END_VAR
  VAR
    r : REF_TO INT;
    rb : REF_TO BA;
    b2 : BA := (i := 10);
    tm : TON;
    rt : REF_TO TON;
    t3 : TON;
    o1 : BG := (n := 3);
    o2 : BG := (n := 6);
    i : IG;
    is : ARRAY [1..2] OF IG;
    pi : REF_TO IG;
  END_VAR
  VAR
    q0 AT %QB0 : SINT;
    q1 AT %QB1 : SINT;
    q2 AT %QB2 : SINT;
    q3 AT %QB3 : SINT;
    q4 AT %QB4 : SINT;
    q5 AT %QB5 : SINT;
    q6 AT %QB6 : SINT;
    q7 AT %QB7 : SINT;
    q8 AT %QB8 : SINT;
    q9 AT %QB9 : SINT;
    q10 AT %QB10 : SINT;
    q11 AT %QB11 : SINT;
    q12 AT %QB12 : SINT;
    q13 AT %QB13 : SINT;
    q14 AT %QB14 : SINT;
    q15 AT %QB15 : SINT;
  END_VAR
  r := Pick(TRUE);
  q0 := INT_TO_SINT(r^);
  Pick(FALSE)^ := 5;
  q1 := INT_TO_SINT(g1);
  IF Nul() = NULL THEN
    q2 := 1;
  END_IF;
  PickP()^.x := 7;
  q3 := INT_TO_SINT(gp.x);
  q4 := INT_TO_SINT(PickP()^.x + 1);
  PickB()^.i := 3;
  PickB()^();
  q5 := INT_TO_SINT(gb.n);
  PickB()^(i := 4);
  q6 := INT_TO_SINT(PickB()^.n);
  rb := REF(gb);
  rb^ := b2;
  gb();
  q7 := INT_TO_SINT(gb.n);
  tm.PT := T#2s;
  IF tm.PT = T#2s THEN
    q8 := 1;
  END_IF;
  rt := REF(gt1);
  rt^.PT := T#3s;
  IF gt1.PT = T#3s THEN
    q9 := 1;
  END_IF;
  PickT()^.PT := T#4s;
  IF gt1.PT = T#4s THEN
    q10 := 1;
  END_IF;
  t3.PT := T#9s;
  rt^ := t3;
  IF gt1.PT = T#9s THEN
    q11 := 1;
  END_IF;
  pi := REF(i);
  pi^ := o1;
  q12 := INT_TO_SINT(i.g());
  pi := REF(is[2]);
  pi^ := o2;
  q13 := INT_TO_SINT(is[2].g());
  IF pi^ <> NULL THEN
    q14 := 1;
  END_IF;
  q15 := INT_TO_SINT(Nul()^);
END_PROGRAM

CONFIGURATION c
  VAR_GLOBAL
    g1 : INT := 1;
    g2 : INT := 2;
    gp : PT;
    gb : BA;
    gt1 : TON;
  END_VAR
  RESOURCE r ON x
    TASK t(INTERVAL := T#10ms, PRIORITY := 1);
    PROGRAM p WITH t : main;
  END_RESOURCE
END_CONFIGURATION

(* ---- refparams.st ---- *)
(* REF_TO as a FUNCTION's and a method's input and output: passed as
   their value, as an interface is (docs/c-output.md §3). Worked by
   hand, i starting at 5, k at 50:

   tick 0. f(r := REF(i), o => p): f is i, 5, then i 6; d not given is
   NULL: 105 (Q0 69 00); p refers to i: 6 (Q2 06 00). b.m(REF(i)): 12
   (Q4 0c 00). f(r := p, d := NULL): i 6, then 7; d NULL: 106 (Q6 6a
   00). b.pick(REF(k), o => p2): k is 50 (Q8 32 00), and p2 refers to
   k, which g bumps through it: 51 (Q10 33 00).
   tick 1: i 7: 107, then 8 (Q0 6b 00, Q2 08 00), m 16 (10 00); 108
   (6c 00), i 9; k 51, then 52 (Q8 33 00, Q10 34 00).
   reference-skip: methods and REF_TO parameters, as `refmore`. *)
FUNCTION f : INT
  VAR_INPUT r : REF_TO INT; d : REF_TO INT; END_VAR
  VAR_OUTPUT o : REF_TO INT; END_VAR
  f := r^;
  r^ := r^ + 1;
  o := r;
  IF d = NULL THEN f := f + 100; END_IF;
END_FUNCTION
FUNCTION g : INT
  VAR_INPUT r : REF_TO INT; END_VAR
  r^ := r^ + 1;
  g := r^;
END_FUNCTION
FUNCTION_BLOCK blk
  METHOD PUBLIC m : INT
    VAR_INPUT r : REF_TO INT; END_VAR
    m := r^ * 2;
  END_METHOD
  METHOD PUBLIC pick : INT
    VAR_INPUT r : REF_TO INT; END_VAR
    VAR_OUTPUT o : REF_TO INT; END_VAR
    pick := r^;
    o := r;
  END_METHOD
END_FUNCTION_BLOCK
PROGRAM main
  VAR i : INT := 5; k : INT := 50; j : INT; p, p2 : REF_TO INT; b : blk; END_VAR
  VAR q AT %QW0 : INT; q2 AT %QW2 : INT; q3 AT %QW4 : INT; q4 AT %QW6 : INT; q5 AT %QW8 : INT; q6 AT %QW10 : INT; END_VAR
  j := f(r := REF(i), o => p);
  q := j;
  q2 := p^;
  q3 := b.m(REF(i));
  q4 := f(r := p, d := NULL);
  q5 := b.pick(r := REF(k), o => p2);
  q6 := g(p2);
END_PROGRAM
CONFIGURATION c RESOURCE r ON PLC TASK t(INTERVAL := T#10ms, PRIORITY := 1); PROGRAM p WITH t : main; END_RESOURCE END_CONFIGURATION

(* ---- refs.st ---- *)
(* References (Ed.3 6.4.4.10): REF_TO an elementary type, through a
   type of its own; to an array element by a computed index, a whole
   array, a structure; REF() and ^ to read, and to write a field or an
   element; = and <> between two references and with NULL; a reference
   as a function block's input, the block reading through it. Each tick
   %IW0 picks what r references: a, b, arr[2], or nothing.
   `r^ := ...` itself is refimage's: the reference compiler's C for it
   does not compile. *)
TYPE
  pair : STRUCT a : INT; b : INT; END_STRUCT;
  rint : REF_TO INT;
  quad : ARRAY[0..3] OF INT;
END_TYPE

FUNCTION_BLOCK bump
VAR_INPUT r : REF_TO INT; inc : INT; END_VAR
VAR_OUTPUT seen : INT; none : BOOL; END_VAR
none := r = NULL;
IF NOT none THEN
  seen := r^ + inc;
END_IF;
END_FUNCTION_BLOCK

PROGRAM main
VAR
  v AT %IW0 : INT;
END_VAR
VAR
  o_a AT %MW0 : INT;
  o_b AT %MW2 : INT;
  o_arr AT %MW4 : INT;
  o_pa AT %MW6 : INT;
  o_pb AT %MW8 : INT;
  o_seen AT %MW10 : INT;
  o_same AT %MX12.0 : BOOL;
  o_null AT %MX12.1 : BOOL;
  o_none AT %MX12.2 : BOOL;
END_VAR
VAR
  a, b, k : INT;
  arr : quad;
  p : pair;
  r, ra : rint;
  rp : REF_TO pair;
  rarr : REF_TO quad;
  f : bump;
  same, isnull : BOOL;
END_VAR
k := v MOD 4;
IF k < 0 THEN
  k := k + 4;
END_IF;
CASE k OF
  0: r := REF(a);
  1: r := REF(b);
  2: r := REF(arr[k]);
ELSE
  r := NULL;
END_CASE;
isnull := r = NULL;
IF r <> NULL THEN
  a := r^ + a + 1;
END_IF;
ra := REF(a);
same := r = ra;
rp := REF(p);
rp^.a := rp^.a + k;
rp^.b := ra^;
rarr := REF(arr);
rarr^[k] := rarr^[k] + 2;
f(r := r, inc := 3);
o_a := a;
o_b := b;
o_arr := arr[2];
o_pa := p.a;
o_pb := p.b;
o_seen := f.seen;
o_same := same;
o_null := isnull;
o_none := f.none;
END_PROGRAM

CONFIGURATION c
  RESOURCE r ON PLC
    TASK t(INTERVAL := T#10ms, PRIORITY := 1);
    PROGRAM inst WITH t : main;
  END_RESOURCE
END_CONFIGURATION

(* ---- refto.st ---- *)
(* CODESYS's REFERENCE TO (the reference-to extension, docs/extensions.md):
   bound with REF= to a variable, to what another one references, to an
   array element by a computed index, to a variable at an address, to a
   structure and to a function block instance; read, written and called
   through without `^`; `.field` and `.output` through it; a function
   block's REFERENCE TO input bound by a call, and kept by a call that does
   not pass it; __ISVALIDREF; REF= 0. At tick 4 %IW0 is 99 and a
   REFERENCE TO unbound by REF= 0 is written: a fault (IECF_FAULT_NULL),
   the statement stores nothing, and the task stops, as at tick 5.
   Worked by hand, a tick at a time: a = vin + 1, p.a = 2a, arr[vin MOD 4]
   (0 if negative) := 7, %QW4 its sum, b grows by vin + 1, %QW6 the sum
   of the vins, %QW0 = a + 100b + p.a: 309, 506, 1118, 1100, then 11400
   before the fault.
   reference-skip: REFERENCE TO is not IEC 61131-3, and the reference
   compiler has none. *)
TYPE pair : STRUCT a : INT; b : BYTE; END_STRUCT; END_TYPE

FUNCTION_BLOCK addto
VAR_INPUT r : REFERENCE TO INT; x : INT; END_VAR
VAR_OUTPUT ok : BOOL; END_VAR
ok := __ISVALIDREF(r);
IF ok THEN r := r + x; END_IF;
END_FUNCTION_BLOCK

FUNCTION_BLOCK acc
VAR_INPUT x : INT; END_VAR
VAR_OUTPUT total : INT; END_VAR
total := total + x;
END_FUNCTION_BLOCK

PROGRAM main
VAR
  vin AT %IW0 : INT;
  q AT %QW0 : INT;
  qb AT %QX2.0 : BOOL;
  qok AT %QX2.1 : BOOL;
  qsum AT %QW4 : INT;
  qtotal AT %QW6 : INT;
END_VAR
VAR
  a, b, i : INT;
  arr : ARRAY[0..3] OF INT;
  p : pair;
  ra, rb, rq : REFERENCE TO INT;
  rp : REFERENCE TO pair;
  f : addto;
  c : acc;
  rc : REFERENCE TO acc;
END_VAR
ra REF= a;
ra := vin;
rb REF= ra;
rb := rb + 1;
rp REF= p;
rp.a := a * 2;
i := vin MOD 4;
IF i < 0 THEN i := 0; END_IF;
ra REF= arr[i];
ra := 7;
rq REF= qsum;
rq := arr[0] + arr[1] + arr[2] + arr[3];
f(r := b, x := vin);
f(x := 1);
qok := f.ok;
rc REF= c;
rc(x := vin);
qtotal := rc.total;
q := a + b * 100 + p.a;
qb := __ISVALIDREF(rb);
rb REF= 0;
IF vin = 99 THEN rb := 5; END_IF;
END_PROGRAM

CONFIGURATION Plant
  RESOURCE r ON PLC
    TASK fast(INTERVAL := T#10ms, PRIORITY := 1);
    PROGRAM p WITH fast : main;
  END_RESOURCE
END_CONFIGURATION

(* ---- replist.st ---- *)
(* A list repeated in an array's initial value (Ed.3 6.4.4.5.2: "A :
   ARRAY[0..5] OF INT := [2(1, 2, 3)] is equivalent to the
   initialization sequence 1, 2, 3, 1, 2, 3"), more values than
   elements ignored (W0008), and a constant's element found in one.
   And two transitions of one chart whose conditions each convert a
   REAL to an integer: a condition left undone is FALSE.
   Worked by hand: c is 1, 2, 3, 1, 2, 3: c[4] 2 (%QB1). K is 4, 5, 6,
   4, 5, 6: K[5] 6 (%QB2). d, five elements of the same list: d[4] 2
   (%QB3). e is [9, 3(2, 7)], four elements: 9, 2, 7, 2: e[3] 2 (%QB4).
   Seq: s0 to s1 when REAL_TO_INT(r) > 2, back when it is > 5; watch
   sets o to s1.X before the transitions are tested (%QB0).
   tick 0: r 3.0: o 0; s0 to s1.         00
   tick 1: o 1; 3 > 5 is not.            01
   tick 2: r 1.0E10: flagged CONVERSION,
           the condition FALSE: s1 stays. 01
   tick 3: r 6.0: o 1; s1 to s0.         01
   tick 4: o 0; s0 to s1.                00
   tick 5: o 1.                          01
   The flag stays from tick 2 on, until the platform clears it.
   reference-skip: the reference compiler's chart tests transitions
   first (sfcdemo), and a conversion out of range is iecf's own. *)
FUNCTION_BLOCK Seq
  VAR_INPUT r : REAL; END_VAR
  VAR_OUTPUT o : INT; END_VAR
  INITIAL_STEP s0 : END_STEP
  TRANSITION FROM s0 TO s1 := REAL_TO_INT(r) > 2; END_TRANSITION
  STEP s1 : END_STEP
  TRANSITION FROM s1 TO s0 := REAL_TO_INT(r) > 5; END_TRANSITION
  INITIAL_STEP w0 : watch(N); END_STEP
  TRANSITION FROM w0 TO w0 := FALSE; END_TRANSITION
  ACTION watch : o := BOOL_TO_INT(s1.X); END_ACTION
END_FUNCTION_BLOCK

PROGRAM main
  VAR CONSTANT K : ARRAY[0..5] OF INT := [2(4, 5, 6)]; END_VAR
  VAR
    c : ARRAY[0..5] OF INT := [2(1, 2, 3)];
    d : ARRAY[0..4] OF INT := [2(1, 2, 3)];
    e : ARRAY[0..3] OF INT := [9, 3(2, 7)];
    s : Seq;
    n : INT;
    r : REAL;
  END_VAR
  VAR
    q0 AT %QB0 : USINT;
    q1 AT %QB1 : USINT;
    q2 AT %QB2 : USINT;
    q3 AT %QB3 : USINT;
    q4 AT %QB4 : USINT;
  END_VAR
  r := 3.0;
  IF n = 2 THEN
    r := 1.0E10;
  ELSIF n > 2 THEN
    r := 6.0;
  END_IF;
  s(r := r);
  q0 := INT_TO_USINT(s.o);
  q1 := INT_TO_USINT(c[4]);
  q2 := INT_TO_USINT(K[5]);
  q3 := INT_TO_USINT(d[4]);
  q4 := INT_TO_USINT(e[3]);
  n := n + 1;
END_PROGRAM
CONFIGURATION c RESOURCE r ON PLC TASK t(INTERVAL := T#10ms, PRIORITY := 1); PROGRAM p WITH t : main; END_RESOURCE END_CONFIGURATION

(* ---- resglobals.st ---- *)
(* The scope of globals (Ed.3 6.5.2.2): each RESOURCE has its own, and
   the configuration's are seen by all. main runs in r1 and in r2, so
   every instance of it, and of the blocks it holds, reaches its own
   resource's g, p, s, a, io, gc, kept: through a pointer the instance
   holds (docs/c-output.md §3). k and shared are the configuration's.
   r1's task runs first (PRIORITY 1), then r2's. Worked by hand:

   tick 0, r1 (g 100): c 101, the VAR_TEMP t 102, arr[1] 103, h.c 104
   (its n 3, lim); h2 := h copies n 3, h2.c 105 (n 6); gc, r1's own
   instance, 106. q 101 + 1000 = 1101 (Q0 4d 04). d.both: bump p.x 11,
   s 'a', 1; a[1] 0 + 1 = 1; inner 107; 1 + 11 = 12 (Q2 0c 00). q3 106
   + readk 1000 = 1106 (Q4 52 04). io 1 (Q20). kept 51 (Q6 33). outp 7
   + 6 = 13 into r1's cout (Q28 0d 00). owner: shared refers to its
   mine.
   r2 (g 200): the same with 201..207: q 1201 (Q10 b1 04); p.x 21, s
   'zza', 3, a[1] 5 + 3 = 8, 29 (Q12 1d 00); q3 1206 (Q14 b6 04); io 1
   (Q21); kept 61 (Q16 3d); outp 9 + 6 = 15 (Q30 0f 00). user: shared^()
   runs r1's instance from r2: it counts r1's g, 108 (Q24 6c 00); mine
   := shared^ copies its values and keeps r2's g: mine() 208 (Q26 d0
   00).
   tick 1, r1 (g 108): c 109, q 1109 (55 04); gc 114, q3 1114 (5a 04);
   p.x 12, s 'aa', a[1] 3, 15; kept 52; h.c n 6, h2 9, outp 16. r2 (g
   208): q 1209, q3 1214, p.x 22, s 'zzaa', a[1] 12, 34; kept 62; outp
   18. user: r1's g 116 (74 00), r2's 216 (d8 00).
   warm, before tick 2: all starts again but kept, RETAIN, each
   resource's own (53, 63), and io, in the image.
   reference-skip: a resource's globals: its C does not link. *)
TYPE
  Pt : STRUCT x : INT; y : INT; END_STRUCT;
  Hold : STRUCT c : counter; n : INT; END_STRUCT;
END_TYPE
FUNCTION_BLOCK counter
  VAR_EXTERNAL g : INT; END_VAR
  VAR_EXTERNAL CONSTANT lim : INT; END_VAR
  VAR_OUTPUT o : INT; n : INT; END_VAR
  g := g + 1;
  n := n + lim;
  o := g;
END_FUNCTION_BLOCK
FUNCTION_BLOCK base
  VAR_EXTERNAL p : Pt; END_VAR
  METHOD PUBLIC bump : INT
    VAR_EXTERNAL s : STRING[8]; END_VAR
    p.x := p.x + 1;
    s := CONCAT(s, 'a');
    bump := LEN(s);
  END_METHOD
END_FUNCTION_BLOCK
FUNCTION_BLOCK derived EXTENDS base
  VAR_EXTERNAL a : ARRAY [0..1] OF INT; END_VAR
  VAR inner : counter; END_VAR
  METHOD PUBLIC both : INT
    a[1] := a[1] + SUPER.bump();
    inner();
    both := a[1] + p.x;
  END_METHOD
END_FUNCTION_BLOCK
FUNCTION readk : INT
  VAR_EXTERNAL k : INT; END_VAR
  readk := k;
END_FUNCTION
PROGRAM main
  VAR_INPUT inp : INT; END_VAR
  VAR_OUTPUT outp : INT; END_VAR
  VAR_EXTERNAL k : INT; io : USINT; gc : counter; kept : USINT; END_VAR
  VAR c : counter; d : derived; arr : ARRAY [0..1] OF counter; h, h2 : Hold; END_VAR
  VAR q AT %Q* : INT; q2 AT %Q* : INT; q3 AT %Q* : INT; q4 AT %Q* : USINT; END_VAR
  VAR_TEMP t : counter; END_VAR
  c();
  t();
  arr[1]();
  h.c();
  h2 := h;
  h2.c();
  gc();
  q := c.o + k;
  q2 := d.both();
  q3 := gc.o + readk();
  io := io + 1;
  kept := kept + 1;
  q4 := kept;
  outp := inp + h2.c.n;
END_PROGRAM
PROGRAM owner
  VAR_EXTERNAL shared : REF_TO counter; END_VAR
  VAR mine : counter; END_VAR
  shared := REF(mine);
END_PROGRAM
PROGRAM user
  VAR_EXTERNAL shared : REF_TO counter; g : INT; END_VAR
  VAR mine : counter; END_VAR
  VAR q AT %QW24 : INT; q2 AT %QW26 : INT; END_VAR
  shared^();
  q := shared^.o;
  mine := shared^;
  mine();
  q2 := mine.o;
END_PROGRAM
CONFIGURATION plant
  VAR_GLOBAL k : INT := 1000; shared : REF_TO counter; END_VAR
  RESOURCE r1 ON PLC
    VAR_GLOBAL g : INT := 100; p : Pt := (x := 10); s : STRING[8]; a : ARRAY [0..1] OF INT; END_VAR
    VAR_GLOBAL io AT %QB20 : USINT; gc : counter; cin : INT := 7; cout AT %QW28 : INT; END_VAR
    VAR_GLOBAL CONSTANT lim : INT := 3; END_VAR
    VAR_GLOBAL RETAIN kept : USINT := 50; END_VAR
    TASK t(INTERVAL := T#10ms, PRIORITY := 1);
    PROGRAM p1 WITH t : main(inp := cin, outp => cout);
    PROGRAM own WITH t : owner;
  END_RESOURCE
  RESOURCE r2 ON PLC
    VAR_GLOBAL g : INT := 200; p : Pt := (x := 20); s : STRING[8] := 'zz'; a : ARRAY [0..1] OF INT := [0, 5]; END_VAR
    VAR_GLOBAL io AT %QB21 : USINT; gc : counter; cin : INT := 9; cout AT %QW30 : INT; END_VAR
    VAR_GLOBAL CONSTANT lim : INT := 3; END_VAR
    VAR_GLOBAL RETAIN kept : USINT := 60; END_VAR
    TASK t(INTERVAL := T#10ms, PRIORITY := 2);
    PROGRAM p1 WITH t : main(inp := cin, outp => cout);
    PROGRAM use WITH t : user;
  END_RESOURCE
  VAR_CONFIG
    r1.p1.q AT %QW0 : INT;
    r1.p1.q2 AT %QW2 : INT;
    r1.p1.q3 AT %QW4 : INT;
    r1.p1.q4 AT %QB6 : USINT;
    r2.p1.q AT %QW10 : INT;
    r2.p1.q2 AT %QW12 : INT;
    r2.p1.q3 AT %QW14 : INT;
    r2.p1.q4 AT %QB16 : USINT;
  END_VAR
END_CONFIGURATION

(* ---- retainloc.st ---- *)
(* RETAIN at an address (Ed.3 Loc_Var_Decls: VAR RETAIN ... AT): its
   initial value is written at a cold start only; at a warm start the
   platform keeps the image bytes, and iecf leaves them (decided
   2026-11-12, florin). Each adds 1 at every tick; a warm restart before
   tick 2. Worked by hand, the M words after set-up, then each tick:
   x RETAIN AT %MW0 := 7:  7, 8, 9 | warm | 10, 11
   y AT %MW2 := 7 (plain): 7, 8, 9 | warm, set again: 7 | 8, 9
   g, a VAR_GLOBAL RETAIN AT %MW4 := 3: 3, 4, 5 | 6, 7
   the block BT's RETAIN z AT %M*, put at %MW6 with 10 by VAR_CONFIG (a
   block's VAR has no full address, Ed.3 Other_Var_Decls): 10, 11, 12
   | 13, 14
   reference-skip: the reference compiler's host makes a warm restart a
   cold one (retain). *)
FUNCTION_BLOCK BT
  VAR RETAIN z AT %M* : INT; END_VAR
  z := z + 1;
END_FUNCTION_BLOCK
PROGRAM main
  VAR RETAIN x AT %MW0 : INT := 7; END_VAR
  VAR y AT %MW2 : INT := 7; END_VAR
  VAR_EXTERNAL g : INT; END_VAR
  VAR b : BT; END_VAR
  x := x + 1;
  y := y + 1;
  g := g + 1;
  b();
END_PROGRAM

CONFIGURATION c
  VAR_GLOBAL RETAIN g AT %MW4 : INT := 3; END_VAR
  RESOURCE r ON x
    TASK t(INTERVAL := T#10ms, PRIORITY := 1);
    PROGRAM p WITH t : main;
  END_RESOURCE
  VAR_CONFIG r.p.b.z AT %MW6 : INT := 10; END_VAR
END_CONFIGURATION

(* ---- retainref.st ---- *)
(* RETAIN references (W0006): kept as they are across a warm restart,
   as CODESYS and TwinCAT keep a pointer in retained memory. Worked by
   hand:

   tick 0: r, a[1] and the global gr are taken, all to x, and n.r to
   n.v; cnt 1. x 1 + 100 + 1000 = 1101 (Q0 4d 04); n.v 10. The blocks h
   and hk each take REF(gx), fresh 1, and count it: gx 2. q2 10 + 2 =
   12 (Q4 0c 00).
   tick 1: x 2202 (9a 08); n.v 20, gx 4: 24 (18 00).
   warm, before tick 2: every reference is RETAIN and still refers to
   what it did; x, n, cnt and gx are RETAIN too. h starts again but for
   its RETAIN r: its fresh is 0 and stays (Q6 00); hk is kept whole
   (Q7 01).
   tick 2: x 3303 (e7 0c), cnt still 1; n.v 30, gx 6: 36 (24 00).
   reference-skip: REF_TO in a structure (its -R); no warm restart. *)
TYPE Node : STRUCT r : REF_TO INT; v : INT; END_STRUCT; END_TYPE
FUNCTION_BLOCK holder
  VAR RETAIN r : REF_TO INT; END_VAR
  VAR_OUTPUT fresh : USINT; END_VAR
  VAR_EXTERNAL gx : INT; END_VAR
  IF r = NULL THEN r := REF(gx); fresh := fresh + 1; END_IF;
  r^ := r^ + 1;
END_FUNCTION_BLOCK
PROGRAM main
  VAR_EXTERNAL gx : INT; gr : REF_TO INT; END_VAR
  VAR RETAIN r : REF_TO INT; x : INT; n : Node; a : ARRAY [0..1] OF REF_TO INT; cnt : USINT; END_VAR
  VAR h : holder; END_VAR
  VAR RETAIN hk : holder; END_VAR
  VAR q AT %QW0 : INT; q1 AT %QB2 : USINT; q2 AT %QW4 : INT; q3 AT %QB6 : USINT; q4 AT %QB7 : USINT; END_VAR
  IF r = NULL THEN
    r := REF(x); n.r := REF(n.v); a[1] := REF(x); gr := REF(x);
    cnt := cnt + 1;
  END_IF;
  r^ := r^ + 1;
  n.r^ := n.r^ + 10;
  a[1]^ := a[1]^ + 100;
  gr^ := gr^ + 1000;
  h();
  hk();
  q := x;
  q1 := cnt;
  q2 := n.v + gx;
  q3 := h.fresh;
  q4 := hk.fresh;
END_PROGRAM
CONFIGURATION plant
  VAR_GLOBAL RETAIN gx : INT; gr : REF_TO INT; END_VAR
  RESOURCE cpu ON PLC
    TASK t(INTERVAL := T#10ms, PRIORITY := 1);
    PROGRAM p WITH t : main;
  END_RESOURCE
END_CONFIGURATION

(* ---- selectdata.st ---- *)
(* SEL, MUX and MOVE of arrays, structures, instances, interfaces and
   references (Ed.3 Table 32, footnote d: allowed for user-defined
   types): the input selected, every input computed first, in order.
   a [1, 2, 3], a2 [4, 5, 6], a3 [7, 8, 9]; b TRUE. Worked by hand:
   SEL(b, a, a2)[1]: 4 (%QB0). SEL(NOT b, a, a2)[2]: 2 (%QB1).
   p.x 7, p2.x 9: SEL(b, p, p2).x 9 (%QB2). MUX(1, a, a2, a3)[3]: 6
   (%QB3); MUX(2, a, a2, a3)[1]: 7 (%QB4). MOVE(a)[2]: 2 (%QB5).
   Sum3(SEL(b, a, a2)), a FUNCTION's input: 4 + 5 + 6, 15 (%QB6).
   f(q := SEL(NOT b, a, a2)), a block's input: f.o[3] 3 (%QB7).
   la AT %MW0, [10, 11, 12]: SEL(b, a, la)[1] 10 (%QB8). Through a
   reference to a2: SEL(b, a, ra^)[2] 5 (%QB9).
   An instance: t2's PT is T#3s; tc := SEL(b, t1, t2) is a copy of t2:
   its PT T#3s (%QB10 1).
   Interfaces: o1 gives 1, o2 2. i := SEL(b, o1, o2): i.g() 2
   (%QB11). j := MUX(0, o1, NULL, i): j.g() 1 (%QB12). k := SEL(b, j,
   NULL) is NULL (%QB13 1).
   References: x1 21, x2 22. r := SEL(b, REF(x1), REF(x2)): r^ 22
   (%QB14). r2 := REF(x1); SEL(b, r, r2)^ := 30 writes x1: 30 (%QB15).
   A FUNCTION's result among them: SEL(b, a, Same(a3))[1] 7 (%QB16).
   Last, MUX(5, a, a2)[1]: K outside 0..1 faults, and the statement
   stores nothing (%QB17 stays 0).
   reference-skip: SEL, MUX, MOVE of arrays and structures, methods:
   the reference compiler refuses them. *)
TYPE
  A3T : ARRAY [1..3] OF INT;
  PT : STRUCT x : INT; y : REAL; END_STRUCT;
END_TYPE
INTERFACE IG
  METHOD g : INT END_METHOD
END_INTERFACE
FUNCTION_BLOCK BG IMPLEMENTS IG
  VAR_INPUT n : INT; END_VAR
  METHOD PUBLIC g : INT
    g := n;
  END_METHOD
END_FUNCTION_BLOCK
FUNCTION Sum3 : INT
  VAR_INPUT q : A3T; END_VAR
  Sum3 := q[1] + q[2] + q[3];
END_FUNCTION
FUNCTION Same : A3T
  VAR_INPUT q : A3T; END_VAR
  Same := q;
END_FUNCTION
FUNCTION_BLOCK FB
  VAR_INPUT q : A3T; END_VAR
  VAR_OUTPUT o : A3T; END_VAR
  o := q;
END_FUNCTION_BLOCK
PROGRAM main
  VAR
    b : BOOL := TRUE;
    a : A3T := [1, 2, 3];
    a2 : A3T := [4, 5, 6];
    a3 : A3T := [7, 8, 9];
    p : PT := (x := 7);
    p2 : PT := (x := 9);
    f : FB;
    ra : REF_TO A3T;
    t1 : TON;
    t2 : TON := (PT := T#3s);
    tc : TON;
    o1 : BG := (n := 1);
    o2 : BG := (n := 2);
    i : IG;
    j : IG;
    k : IG;
    x1 : INT := 21;
    x2 : INT := 22;
    r : REF_TO INT;
    r2 : REF_TO INT;
    v5 : INT := 5;
  END_VAR
  VAR
    la AT %MW0 : A3T := [10, 11, 12];
  END_VAR
  VAR
    q0 AT %QB0 : SINT;
    q1 AT %QB1 : SINT;
    q2 AT %QB2 : SINT;
    q3 AT %QB3 : SINT;
    q4 AT %QB4 : SINT;
    q5 AT %QB5 : SINT;
    q6 AT %QB6 : SINT;
    q7 AT %QB7 : SINT;
    q8 AT %QB8 : SINT;
    q9 AT %QB9 : SINT;
    q10 AT %QB10 : SINT;
    q11 AT %QB11 : SINT;
    q12 AT %QB12 : SINT;
    q13 AT %QB13 : SINT;
    q14 AT %QB14 : SINT;
    q15 AT %QB15 : SINT;
    q16 AT %QB16 : SINT;
    q17 AT %QB17 : SINT;
  END_VAR
  q0 := INT_TO_SINT(SEL(b, a, a2)[1]);
  q1 := INT_TO_SINT(SEL(NOT b, a, a2)[2]);
  q2 := INT_TO_SINT(SEL(b, p, p2).x);
  q3 := INT_TO_SINT(MUX(1, a, a2, a3)[3]);
  q4 := INT_TO_SINT(MUX(2, a, a2, a3)[1]);
  q5 := INT_TO_SINT(MOVE(a)[2]);
  q6 := INT_TO_SINT(Sum3(SEL(b, a, a2)));
  f(q := SEL(NOT b, a, a2));
  q7 := INT_TO_SINT(f.o[3]);
  q8 := INT_TO_SINT(SEL(b, a, la)[1]);
  ra := REF(a2);
  q9 := INT_TO_SINT(SEL(b, a, ra^)[2]);
  tc := SEL(b, t1, t2);
  IF tc.PT = T#3s THEN
    q10 := 1;
  END_IF;
  i := SEL(b, o1, o2);
  q11 := INT_TO_SINT(i.g());
  j := MUX(0, o1, NULL, i);
  q12 := INT_TO_SINT(j.g());
  k := SEL(b, j, NULL);
  IF k = NULL THEN
    q13 := 1;
  END_IF;
  r := SEL(b, REF(x1), REF(x2));
  q14 := INT_TO_SINT(r^);
  r2 := REF(x1);
  SEL(b, r, r2)^ := 30;
  q15 := INT_TO_SINT(x1);
  q16 := INT_TO_SINT(SEL(b, a, Same(a3))[1]);
  q17 := INT_TO_SINT(MUX(v5, a, a2)[1]);
END_PROGRAM

CONFIGURATION c
  RESOURCE r ON x
    TASK t(INTERVAL := T#10ms, PRIORITY := 1);
    PROGRAM p WITH t : main;
  END_RESOURCE
END_CONFIGURATION

(* ---- seqpath.st ---- *)
(* An element of an in-out array passed to a FUNCTION that writes a
   global: the call is sequenced (its operands each on a line, as it may
   change what they read), and the element's index is found once. Until
   2026-11-19 it was found twice, the first line left unused, which C's
   -Wall -Werror refused (found in the OSCAT BASIC library's HOLIDAY).
   Worked by hand: hs[1].d is 5; G(y, hs[i].d) with y 0 is 5, gx 1
   (%QW2); 5 = y fails on the first tick: y := y + hs[i].d, 5 (%QW0);
   the second tick G(5, 5) = 10, gx 2; 10 = 5 fails, y := 10. *)
TYPE H : STRUCT d : INT; END_STRUCT; END_TYPE

FUNCTION G : INT
  VAR_INPUT a, b : INT; END_VAR
  VAR_EXTERNAL gx : INT; END_VAR
  gx := gx + 1;
  G := a + b;
END_FUNCTION

FUNCTION_BLOCK FB
  VAR_IN_OUT hs : ARRAY[0..3] OF H; END_VAR
  VAR_OUTPUT y : INT; END_VAR
  VAR i : INT := 1; END_VAR
  IF G(y, hs[i].d) = y THEN
    y := -1;
  ELSE
    y := y + hs[i].d;
  END_IF;
END_FUNCTION_BLOCK

PROGRAM main
  VAR a : ARRAY[0..3] OF H := [(d := 0), (d := 5)]; f : FB; END_VAR
  VAR_EXTERNAL gx : INT; END_VAR
  VAR q0 AT %QW0 : INT; q1 AT %QW2 : INT; END_VAR
  f(hs := a);
  q0 := f.y;
  q1 := gx;
END_PROGRAM

CONFIGURATION cf
  VAR_GLOBAL gx : INT; END_VAR
  RESOURCE r ON x
    TASK tk(INTERVAL := T#10ms, PRIORITY := 1);
    PROGRAM p WITH tk : main;
  END_RESOURCE
END_CONFIGURATION

(* ---- shadow.st ---- *)
(* A global named as one further out hides it where it is seen (as a
   local name does in CODESYS; Ed.3 gives no rule): r1's g hides the
   configuration's in r1, the PROGRAM own's g hides r1's for what own
   holds, and r2, which declares none, sees the configuration's.
   Worked by hand:

   tick 0. r1.a (main): the block counts r1's g, 100 + 1 = 101; main
   adds 10: 111 (Q0 6f 00). r1.b (own): its block counts own's g, 1000
   + 1 = 1001, own adds 100: 1101 (Q2 4d 04). r2.a (main): the
   configuration's g, 1 + 1 + 10 = 12 (Q4 0c 00). r1.a's connection i
   := g reads r1's g before a runs, 100, and o => res puts it in r1's
   res (Q6 64 00).
   tick 1: 122 (7a 00), 1202 (b2 04), 23 (17 00), res 111 (6f 00).
   reference-skip: a global named as an outer one: the reference
   compiler refuses it. *)
FUNCTION_BLOCK counter
  VAR_EXTERNAL g : INT; END_VAR
  g := g + 1;
END_FUNCTION_BLOCK
PROGRAM main
  VAR_INPUT i : INT; END_VAR
  VAR_OUTPUT o : INT; END_VAR
  VAR_EXTERNAL g : INT; END_VAR
  VAR c : counter; END_VAR
  VAR q AT %Q* : INT; END_VAR
  c();
  g := g + 10;
  q := g;
  o := i;
END_PROGRAM
PROGRAM own
  VAR_GLOBAL g : INT := 1000; END_VAR
  VAR c : counter; END_VAR
  VAR q AT %QW2 : INT; END_VAR
  c();
  g := g + 100;
  q := g;
END_PROGRAM
CONFIGURATION plant
  VAR_GLOBAL g : INT := 1; END_VAR
  RESOURCE r1 ON PLC
    VAR_GLOBAL g : INT := 100; END_VAR
    VAR_GLOBAL res AT %QW6 : INT; END_VAR
    TASK t(INTERVAL := T#10ms, PRIORITY := 1);
    PROGRAM a WITH t : main(i := g, o => res);
    PROGRAM b WITH t : own;
  END_RESOURCE
  RESOURCE r2 ON PLC
    TASK t(INTERVAL := T#10ms, PRIORITY := 2);
    PROGRAM a WITH t : main;
  END_RESOURCE
  VAR_CONFIG
    r1.a.q AT %QW0 : INT;
    r2.a.q AT %QW4 : INT;
  END_VAR
END_CONFIGURATION

(* ---- shadowing.st ---- *)
(* shadowing: a POU's variable named as a type, a POU or a standard
   block or function; in its POU the name is the variable. Worked by
   hand:
   Length, a FUNCTION_BLOCK, counts its calls in n; Speed, a TYPE, a
   structure. In main: length : INT (the block's name) := 7; speed :
   Speed, a variable of the type it is named as, speed.v := 3; tp : BOOL
   (TP, a standard block) beside t : TP, an instance of the block, which
   the name still means as a type; max : INT := 40 (MAX, a standard
   function).
   %QB0: length + speed.v, 10. %QB1: c, an instance of Length, called
   twice: its n is 2. %QB2: t's Q, TRUE on its first call (PT T#1s),
   copied into tp: 1. %QB3: max + 2, 42.
   reference-skip: shadowing is CODESYS's, not IEC 61131-3. *)
FUNCTION_BLOCK Length
  VAR_OUTPUT n : INT; END_VAR
  n := n + 1;
END_FUNCTION_BLOCK

TYPE Speed : STRUCT v : INT; END_STRUCT; END_TYPE

PROGRAM main
  VAR
    length : INT := 7;
    speed : Speed;
    c : Length;
    tp : BOOL;
    t : TP;
    max : INT := 40;
  END_VAR
  VAR
    q0 AT %QB0 : SINT;
    q1 AT %QB1 : SINT;
    q2 AT %QB2 : SINT;
    q3 AT %QB3 : SINT;
  END_VAR
  speed.v := 3;
  q0 := INT_TO_SINT(length + speed.v);
  c();
  c();
  q1 := INT_TO_SINT(c.n);
  t(IN := TRUE, PT := T#1s);
  tp := t.Q;
  q2 := SEL(tp, SINT#0, SINT#1);
  q3 := INT_TO_SINT(max + 2);
END_PROGRAM

CONFIGURATION cf
  RESOURCE r ON x
    TASK tk(INTERVAL := T#10ms, PRIORITY := 1);
    PROGRAM p WITH tk : main;
  END_RESOURCE
END_CONFIGURATION

(* ---- starinout.st ---- *)
(* A structure with `*` components given to an in-out (Ed.3 6.4.4.8,
   6.5.5.4): the in-out holds no data of its own, it binds the caller's
   variable, whose components VAR_CONFIG places. A FUNCTION_BLOCK and a
   FUNCTION each reach the image through it.
   Worked by hand, each tick: d.a := d.a + 10 (a at %MW0, from 0);
   r(x := d) sets q (%QW0) to a + 1; Twice(x := d) sets o (%QW2) to
   a * 2 and gives it, into %QW4.
   Tick 1: a 10, q 11, o 20, 20. Tick 2: a 20, q 21, o 40, 40.
   reference-skip: VAR_CONFIG, as varconfig. *)
TYPE Io : STRUCT
  a AT %M* : INT;
  q AT %Q* : INT;
  o AT %Q* : INT;
END_STRUCT;
END_TYPE

FUNCTION_BLOCK Robot
  VAR_IN_OUT x : Io; END_VAR
  x.q := x.a + 1;
END_FUNCTION_BLOCK

FUNCTION Twice : INT
  VAR_IN_OUT x : Io; END_VAR
  x.o := x.a * 2;
  Twice := x.o;
END_FUNCTION

PROGRAM main
  VAR d : Io; END_VAR
  VAR r : Robot; END_VAR
  VAR t AT %QW4 : INT; END_VAR
  d.a := d.a + 10;
  r(x := d);
  t := Twice(x := d);
END_PROGRAM

CONFIGURATION cf
  RESOURCE rs ON x
    TASK tk(INTERVAL := T#10ms, PRIORITY := 1);
    PROGRAM p WITH tk : main;
  END_RESOURCE
  VAR_CONFIG
    rs.p.d.a AT %MW0 : INT;
    rs.p.d.q AT %QW0 : INT;
    rs.p.d.o AT %QW2 : INT;
  END_VAR
END_CONFIGURATION

(* ---- stdinout.st ---- *)
(* A standard function block's instance as a VAR_IN_OUT: the caller's
   own instance, by its address, in a FUNCTION, in one that passes it
   on, and in a FUNCTION_BLOCK; given a variable, an array's element
   and what a reference refers to.
   tick is TRUE at ticks 0, 2, 4. Count calls c(CU := up, PV := 3).
   Count(c1, tick): c1 counts the three rising edges: 1 1 2 2 3 3
   (%QB0), and c1.Q, CV >= 3, is TRUE at ticks 4 and 5 (%QX4.0).
   Pass(cs[2], tick) gives it to Count: the same, 1 1 2 2 3 3 (%QB1),
   and it is cs[2] that counted (%QB5).
   Count(r^, TRUE), r referring to cs[1]: one rising edge, 1 at every
   tick (%QB2).
   Hold runs the TON it is given, PT 20 ms, the interval 10 ms: IN TRUE
   from tick 0, Q at tick 2 (%QX3.0), and it is t1 that ran (%QX6.0).
   reference-skip: a block instance as an in-out: iec2c crashes. *)
FUNCTION Count : INT
  VAR_IN_OUT c : CTU; END_VAR
  VAR_INPUT up : BOOL; END_VAR
  c(CU := up, PV := 3);
  Count := c.CV;
END_FUNCTION
FUNCTION Pass : INT
  VAR_IN_OUT c : CTU; END_VAR
  VAR_INPUT up : BOOL; END_VAR
  Pass := Count(c, up);
END_FUNCTION
FUNCTION_BLOCK Hold
  VAR_IN_OUT tm : TON; END_VAR
  VAR_INPUT go : BOOL; END_VAR
  VAR_OUTPUT q : BOOL; END_VAR
  tm(IN := go, PT := T#20ms);
  q := tm.Q;
END_FUNCTION_BLOCK
PROGRAM main
  VAR
    c1 : CTU;
    cs : ARRAY [1..2] OF CTU;
    t1 : TON;
    h : Hold;
    r : REF_TO CTU;
    tick : BOOL;
  END_VAR
  VAR
    q0 AT %QB0 : SINT;
    q1 AT %QB1 : SINT;
    q2 AT %QB2 : SINT;
    q3 AT %QX3.0 : BOOL;
    q4 AT %QX4.0 : BOOL;
    q5 AT %QB5 : SINT;
    q6 AT %QX6.0 : BOOL;
  END_VAR
  tick := NOT tick;
  q0 := INT_TO_SINT(Count(c1, tick));
  q1 := INT_TO_SINT(Pass(cs[2], tick));
  r := REF(cs[1]);
  q2 := INT_TO_SINT(Count(r^, TRUE));
  h(tm := t1, go := TRUE);
  q3 := h.q;
  q4 := c1.Q;
  q5 := INT_TO_SINT(cs[2].CV);
  q6 := t1.Q;
END_PROGRAM

CONFIGURATION c
  RESOURCE r ON x
    TASK t(INTERVAL := T#10ms, PRIORITY := 1);
    PROGRAM p WITH t : main;
  END_RESOURCE
END_CONFIGURATION

(* ---- subparams.st ---- *)
(* A subrange as a FUNCTION's input, output, in-out and result, and as
   a FUNCTION_BLOCK's in-out; and what a subrange starts as: its lower
   limit (Ed.3 6.4.4.4.2), unless its type or declaration says.
   SRT is INT (2..5); S3 is INT (2..5) := 4. Worked by hand, the same
   at every tick:
   x : INT (1..5), y : SRT, z : S3, a : ARRAY OF SRT start as 1, 2, 4,
   2: x + y + z + a[2] is 9 (%QB0).
   Sum(p : INT (0..5), q : SRT, z : S3 := 3) adds them. Sum(), each
   input its initial value, 0 + 2 + 3: 5 (%QB1). Sum(1, 3, 4): 8 (%QB2).
   Res : SRT, set only when x > 0: Res(0) is its lower limit, 2 (%QB3);
   Res(4): 4 (%QB4).
   Out(x, o => s) sets its output o : SRT to x and gives it: with 3, 3
   (%QB5), and s is 3 (%QB6).
   From here a value is outside its subrange: clamped to the bound it
   passed and flagged CONVERSION, first at the call that gives Sum's
   input p 9, Sum(9, 3, 4) at line 91: 5 + 3 + 4, 12 (%QB7). Res(9): 5 (%QB8).
   Out(1, o => s): 2 (%QB9), and s is 2 (%QB10).
   An in-out is the caller's variable, a store through it clamped to
   the in-out's bounds: s := 4; Bump(s) adds 10, 5 (%QB11), and s is 5
   (%QB12). The block Hold takes 10 from its in-out: h(io := s) leaves
   s 2 (%QB13). n, an INT, given to Bump: n := 4 becomes 5 (%QB14,
   %QB15).
   reference-skip: a call with no arguments: refused; and a subrange
   starts at 0 there (Ed.3 6.4.4.4: its lower limit), not clamped into
   one. *)
TYPE
  SRT : INT (2..5);
  S3 : INT (2..5) := 4;
END_TYPE
FUNCTION Sum : INT
  VAR_INPUT p : INT (0..5); q : SRT; z : S3 := 3; END_VAR
  Sum := p + q + z;
END_FUNCTION
FUNCTION Res : SRT
  VAR_INPUT x : INT; END_VAR
  IF x > 0 THEN
    Res := x;
  END_IF;
END_FUNCTION
FUNCTION Out : INT
  VAR_INPUT x : INT; END_VAR
  VAR_OUTPUT o : SRT; END_VAR
  o := x;
  Out := o;
END_FUNCTION
FUNCTION Bump : INT
  VAR_IN_OUT io : SRT; END_VAR
  io := io + 10;
  Bump := io;
END_FUNCTION
FUNCTION_BLOCK Hold
  VAR_IN_OUT io : SRT; END_VAR
  io := io - 10;
END_FUNCTION_BLOCK
PROGRAM main
  VAR
    x : INT (1..5);
    y : SRT;
    z : S3;
    a : ARRAY [1..2] OF SRT;
    s : SRT;
    n : INT;
    h : Hold;
  END_VAR
  VAR
    q0 AT %QB0 : SINT;
    q1 AT %QB1 : SINT;
    q2 AT %QB2 : SINT;
    q3 AT %QB3 : SINT;
    q4 AT %QB4 : SINT;
    q5 AT %QB5 : SINT;
    q6 AT %QB6 : SINT;
    q7 AT %QB7 : SINT;
    q8 AT %QB8 : SINT;
    q9 AT %QB9 : SINT;
    q10 AT %QB10 : SINT;
    q11 AT %QB11 : SINT;
    q12 AT %QB12 : SINT;
    q13 AT %QB13 : SINT;
    q14 AT %QB14 : SINT;
    q15 AT %QB15 : SINT;
  END_VAR
  q0 := INT_TO_SINT(x + y + z + a[2]);
  q1 := INT_TO_SINT(Sum());
  q2 := INT_TO_SINT(Sum(1, 3, 4));
  q3 := INT_TO_SINT(Res(0));
  q4 := INT_TO_SINT(Res(4));
  n := 3;
  q5 := INT_TO_SINT(Out(x := n, o => s));
  q6 := INT_TO_SINT(s);
  q7 := INT_TO_SINT(Sum(9, 3, 4));
  q8 := INT_TO_SINT(Res(9));
  q9 := INT_TO_SINT(Out(x := 1, o => s));
  q10 := INT_TO_SINT(s);
  s := 4;
  q11 := INT_TO_SINT(Bump(s));
  q12 := INT_TO_SINT(s);
  h(io := s);
  q13 := INT_TO_SINT(s);
  n := 4;
  q14 := INT_TO_SINT(Bump(n));
  q15 := INT_TO_SINT(n);
END_PROGRAM

CONFIGURATION c
  RESOURCE r ON x
    TASK t(INTERVAL := T#10ms, PRIORITY := 1);
    PROGRAM p WITH t : main;
  END_RESOURCE
END_CONFIGURATION

(* ---- subrange.st ---- *)
(* A value stored into a subrange outside its bounds is clamped to the
   bound it passed and flagged (docs/dependencies.md, decided
   2026-11-06): by an assignment, into an array's element and a
   structure's field, into a function block's input; a FOR over a
   subrange stops at the bound it would pass. At tick 1, 150 leaves
   percent: p is 100, and the FOR to 150 stops at 3; at tick 2, -5: p is
   0, and the FOR to -5 does not run. The first is flagged, code 4 at
   line 41. The reference compiler stores unchecked but at the function block's input,
   and its FOR leaves the subrange; iecf's trace is
   subrange.iecf.trace. *)
TYPE
  percent : INT (0..100) := 50;
  pair : STRUCT
    a : percent;
  END_STRUCT;
END_TYPE

FUNCTION_BLOCK hold
VAR_INPUT v : percent; END_VAR
VAR_OUTPUT o : INT; END_VAR
o := v;
END_FUNCTION_BLOCK

PROGRAM main
VAR
  k AT %IW0 : INT;
  r_p AT %MW0 : INT;
  r_arr AT %MW2 : INT;
  r_pair AT %MW4 : INT;
  r_fb AT %MW6 : INT;
  r_for AT %MW8 : INT;
END_VAR
VAR
  p : percent;
  arr : ARRAY [1..2] OF percent;
  pr : pair;
  h : hold;
  i : INT (1..3);
  n : INT;
END_VAR
p := k;
arr[2] := k * 2;
pr.a := k + 1;
h(v := k - 1);
r_p := p;
r_arr := arr[2];
r_pair := pr.a;
r_fb := h.o;
n := 0;
FOR i := 1 TO k DO
  n := n + 1;
END_FOR;
r_for := n;
END_PROGRAM

CONFIGURATION plant
  RESOURCE r ON PLC
    TASK fast(INTERVAL := T#10ms, PRIORITY := 0);
    PROGRAM p WITH fast : main;
  END_RESOURCE
END_CONFIGURATION

(* ---- temp.st ---- *)
(* VAR_TEMP (Ed.3 6.5.2.2): set to its initial value at each call of its
   PROGRAM or FUNCTION_BLOCK, where VAR keeps its value. The reference compiler reads
   Ed.2, where VAR_TEMP takes no initial value: each starts at 0. An
   array in VAR_TEMP is left out: the reference compiler's C for it does not compile
   (PROPOSAL.md §1b). *)
FUNCTION_BLOCK acc
VAR_INPUT x : INT; END_VAR
VAR_OUTPUT kept, fresh : INT; END_VAR
VAR total : INT; END_VAR
VAR_TEMP part : INT; END_VAR
total := total + x;
part := part + x;
kept := total;
fresh := part;
END_FUNCTION_BLOCK

PROGRAM main
VAR
  k AT %IW0 : INT;
  r_kept AT %MW0 : INT;
  r_fresh AT %MW2 : INT;
  r_tmp AT %MW4 : INT;
END_VAR
VAR
  a : acc;
END_VAR
VAR_TEMP
  tmp : INT;
  flag : BOOL;
END_VAR
a(x := k);
tmp := tmp + k;
flag := NOT flag;
r_kept := a.kept;
r_fresh := a.fresh;
IF flag THEN r_tmp := tmp; END_IF;
END_PROGRAM

CONFIGURATION plant
  RESOURCE r ON PLC
    TASK fast(INTERVAL := T#10ms, PRIORITY := 0);
    PROGRAM p WITH fast : main;
  END_RESOURCE
END_CONFIGURATION

(* ---- timefunc.st ---- *)
(* TIME() (the time-function extension): the running task's clock, in
   milliseconds. The task runs every 10 ms, its clock 0, 10, 20, 30 ms on
   ticks 0..3. Worked by hand:
   %QB0: TIME() in the PROGRAM, as ms / 10: 0, 1, 2, 3.
   %QB1: Now10, a FUNCTION reading it too: the same.
   %QB2: Since, a block that keeps its first reading, OSCAT's way of
   measuring (T_PLC_MS): TIME() - start, 0, 10, 20, 30 ms, / 10.
   %QX3.0: a TON of PT T#25ms beside it, started on tick 0: Q from
   tick 3 (30 ms) on, as Since passes 25 ms.
   reference-skip: TIME() is CODESYS's, not IEC 61131-3. *)
FUNCTION Now10 : SINT
  Now10 := DINT_TO_SINT(TIME_TO_DINT(TIME()) / 10);
END_FUNCTION

FUNCTION_BLOCK Since
  VAR_OUTPUT elapsed : TIME; END_VAR
  VAR start : TIME; first : BOOL := TRUE; END_VAR
  IF first THEN
    start := TIME();
    first := FALSE;
  END_IF;
  elapsed := TIME() - start;
END_FUNCTION_BLOCK

PROGRAM main
  VAR s : Since; t : TON; END_VAR
  VAR
    q0 AT %QB0 : SINT;
    q1 AT %QB1 : SINT;
    q2 AT %QB2 : SINT;
    q3 AT %QX3.0 : BOOL;
  END_VAR
  q0 := DINT_TO_SINT(TIME_TO_DINT(TIME()) / 10);
  q1 := Now10();
  s();
  q2 := DINT_TO_SINT(TIME_TO_DINT(s.elapsed) / 10);
  t(IN := TRUE, PT := T#25ms);
  q3 := t.Q;
END_PROGRAM

CONFIGURATION cf
  RESOURCE r ON x
    TASK tk(INTERVAL := T#10ms, PRIORITY := 1);
    PROGRAM p WITH tk : main;
  END_RESOURCE
END_CONFIGURATION

(* ---- toplist.st ---- *)
(* A VAR_GLOBAL list outside any CONFIGURATION, as CODESYS writes one:
   seen by every configuration, each with its own of each variable; the
   configuration's own lim hides the list's. A plain, a CONSTANT, a
   RETAIN and a located one, reached by a program and a block. Worked
   by hand:

   tick 0: the block adds the list's kk, 4, to its g: 9; q is g + the
   configuration's lim, 100: 109 (Q0 6d 00); kept 11 (Q2); out 1 (Q6).
   tick 1: g 13, 113 (71 00); kept 12; out 2.
   warm, before tick 2: g 5 again; kept, RETAIN, stays; out is in the
   image.
   tick 2: 109; kept 13; out 3.
   reference-skip: the reference compiler has no VAR_GLOBAL outside a
   CONFIGURATION. *)
VAR_GLOBAL g : INT := 5; lim : INT := 3; END_VAR
VAR_GLOBAL CONSTANT kk : INT := 4; END_VAR
VAR_GLOBAL RETAIN kept : INT := 10; out AT %QW6 : INT; END_VAR
FUNCTION_BLOCK counter
  VAR_EXTERNAL g : INT; END_VAR
  VAR_EXTERNAL CONSTANT kk : INT; END_VAR
  g := g + kk;
END_FUNCTION_BLOCK
PROGRAM main
  VAR_EXTERNAL g : INT; lim : INT; kept : INT; out : INT; END_VAR
  VAR c : counter; END_VAR
  VAR q AT %Q* : INT; q2 AT %Q* : INT; END_VAR
  c();
  kept := kept + 1;
  q := g + lim;
  q2 := kept;
  out := out + 1;
END_PROGRAM
CONFIGURATION A
  VAR_GLOBAL lim : INT := 100; END_VAR
  RESOURCE r1 ON PLC TASK t(INTERVAL := T#10ms, PRIORITY := 1); PROGRAM p WITH t : main; END_RESOURCE
  VAR_CONFIG r1.p.q AT %QW0 : INT; r1.p.q2 AT %QW2 : INT; END_VAR
END_CONFIGURATION

(* ---- underscorenames.st ---- *)
(* Names starting with one underscore (Ed.3 6.1.2 allows it), in a
   namespace: iecf keys LIB._BASE as LIB___BASE and a method as its
   type's key, `__` and its name, so the namespace and the type are
   found at the `__` before the underscore. INTERNAL called from a type
   of the namespace, a method's input given the type's constant, an
   override called through THIS, SUPER, a REF_TO the base, and a method
   through an interface.
   Worked by hand, one tick: d._Run(): THIS._Bump() is _DERIVED's, amount
   := _k 5, SUPER._Bump(amount := 6): n 6; THIS._Close() n 12.
   b._Bump(): amount 5, b.n 5. r := REF(d); r^._Bump(): _DERIVED's: d.n 18.
   i := d; i._Get() 18.
   %QW0 18, %QW2 5, %QW4 18.
   reference-skip: NAMESPACE, METHOD, INTERFACE are Ed.3's; the
   reference compiler (Ed.2) has none. *)
NAMESPACE Lib
  INTERFACE _Itf
    METHOD _Get : INT
    END_METHOD
  END_INTERFACE

  FUNCTION_BLOCK _Base
    VAR CONSTANT _k : INT := 5; END_VAR
    VAR_OUTPUT n : INT; END_VAR
    METHOD PUBLIC _Bump
      VAR_INPUT amount : INT := _k; END_VAR
      n := n + amount;
    END_METHOD
    METHOD INTERNAL _Close
      n := n * 2;
    END_METHOD
  END_FUNCTION_BLOCK

  FUNCTION_BLOCK _Derived EXTENDS _Base IMPLEMENTS _Itf
    METHOD PUBLIC OVERRIDE _Bump
      VAR_INPUT amount : INT := _k; END_VAR
      SUPER._Bump(amount := amount + 1);
    END_METHOD
    METHOD PUBLIC _Get : INT
      _Get := n;
    END_METHOD
    METHOD PUBLIC _Run
      THIS._Bump();
      THIS._Close();
    END_METHOD
  END_FUNCTION_BLOCK
END_NAMESPACE

PROGRAM main
  VAR
    d : Lib._Derived; b : Lib._Base; r : REF_TO Lib._Base; i : Lib._Itf;
  END_VAR
  VAR
    q0 AT %QW0 : INT; q1 AT %QW2 : INT; q2 AT %QW4 : INT;
  END_VAR
  d._Run();
  b._Bump();
  r := REF(d);
  r^._Bump();
  i := d;
  q0 := i._Get();
  q1 := b.n;
  q2 := d.n;
END_PROGRAM

CONFIGURATION cf
  RESOURCE r ON x
    TASK tk(INTERVAL := T#10ms, PRIORITY := 1);
    PROGRAM p WITH tk : main;
  END_RESOURCE
END_CONFIGURATION

(* ---- undonecalls.st ---- *)
(* A real that does not fit its integer, in the index of a place a call
   takes: the statement is left undone (docs/behaviour/conversions.md).
   A FUNCTION after the conversion is not called, a block is not called,
   and nothing is stored - not into the element the placeholder, 0,
   would find. r is 1.0E10, beyond INT; r2 3.0. Worked by hand, the
   same each tick but the counts:
   n := Two(o => a[REAL_TO_INT(r)]): an output's place is found after
   the call, so Two is called (calls 1) and neither a[0] nor n stored.
   n := Inc(a[REAL_TO_INT(r) + 1]): Inc not called, a[1] 0, n 7.
   n := Two(i := REAL_TO_INT(r), o => x): not called, x and n kept.
   n := REAL_TO_INT(r) + Inc(a[2]): not called, a[2] 0.
   Two(o => a[REAL_TO_INT(r)]), a statement: called (calls 2), not
   stored. SPLIT_DATE into a[REAL_TO_INT(r)] and a[1]: neither stored.
   The block calls not made, the index in a place found before the
   block runs: an instance by it; an in-out by it, alone and with EN,
   whose ENO then keeps bs[1] TRUE; an array in-out; an instance
   in-out. Those whose index is where an output goes - an output, a
   STRING output, ENO, TON's Q into bs[..] - are made, the place found
   after the block runs, as a FUNCTION's output's is, and not stored.
   So f runs three times there (f.q 3, x 3); then
   f(q => a[REAL_TO_INT(r2)]): f.q 4 into a[3]; f(): f.q 5, x 5. The
   next tick each again: f.q 10, x 10, a[3] 9.
   %QB0 a[0] 0, %QB1 a[1] 0, %QB2 a[2] 0, %QB3 n 7, %QB4 calls 2 then
   4, %QB5 f.q 5 then 10, %QB6 x 5 then 10, %QB7 fs[0].q 0, %QB8 g.n +
   u.n 0, %QB9 a[3] 4 then 9; %QX10.0 bs[0] TRUE, %QX10.1 bs[1] TRUE,
   %QX10.2 ss[0] still '', %QX10.3 tm.Q TRUE (PT 0s, called once).
   And the same index in a whole value read, in an instance whose
   input is set, in REF(): row := aa[REAL_TO_INT(r)] keeps row[0] 5
   (%QB11); fs[REAL_TO_INT(r)].d := 9 leaves fs[0].d 0 (%QB12);
   rf := REF(a[REAL_TO_INT(r)]) leaves rf NULL (%QX10.4).
   Flagged CONVERSION at the first, no fault.
   reference-skip: a statement left undone is iecf's own. *)
FUNCTION Inc : INT
  VAR_IN_OUT c : INT; END_VAR
  c := c + 1;
  Inc := c;
END_FUNCTION

FUNCTION Two : INT
  VAR_INPUT i : INT; END_VAR
  VAR_OUTPUT o : INT; END_VAR
  VAR_EXTERNAL calls : INT; END_VAR
  calls := calls + 1;
  o := 2 + i;
  Two := 1;
END_FUNCTION

FUNCTION_BLOCK Cnt
  VAR_INPUT d : INT; END_VAR
  VAR_IN_OUT c : INT; END_VAR
  VAR_OUTPUT q : INT; s : STRING[4]; END_VAR
  q := q + 1;
  c := c + d;
  s := 'ab';
END_FUNCTION_BLOCK

FUNCTION_BLOCK Arr
  VAR_IN_OUT v : ARRAY[0..1] OF INT; END_VAR
  VAR_OUTPUT n : INT; END_VAR
  n := n + 1;
  v[0] := v[0] + 1;
END_FUNCTION_BLOCK

FUNCTION_BLOCK Use
  VAR_IN_OUT f : Cnt; END_VAR
  VAR_OUTPUT n : INT; END_VAR
  n := n + 1;
END_FUNCTION_BLOCK

PROGRAM main
  VAR_EXTERNAL calls : INT; END_VAR
  VAR
    a : ARRAY[0..3] OF INT;
    aa : ARRAY[0..1] OF ARRAY[0..1] OF INT;
    ss : ARRAY[0..1] OF STRING[4];
    bs : ARRAY[0..3] OF BOOL := [4(TRUE)];
    r : REAL := 1.0E10;
    r2 : REAL := 3.0;
    x : INT;
    n : INT := 7;
    f : Cnt;
    fs : ARRAY[0..1] OF Cnt;
    g : Arr;
    u : Use;
    tm : TON;
    row : ARRAY[0..1] OF INT := [5, 6];
    rf : REF_TO INT;
  END_VAR
  VAR
    q0 AT %QB0 : SINT;
    q1 AT %QB1 : SINT;
    q2 AT %QB2 : SINT;
    q3 AT %QB3 : SINT;
    q4 AT %QB4 : SINT;
    q5 AT %QB5 : SINT;
    q6 AT %QB6 : SINT;
    q7 AT %QB7 : SINT;
    q8 AT %QB8 : SINT;
    q9 AT %QB9 : SINT;
    b0 AT %QX10.0 : BOOL;
    b1 AT %QX10.1 : BOOL;
    b2 AT %QX10.2 : BOOL;
    b3 AT %QX10.3 : BOOL;
    b4 AT %QX10.4 : BOOL;
    q11 AT %QB11 : SINT;
    q12 AT %QB12 : SINT;
  END_VAR
  n := Two(o => a[REAL_TO_INT(r)]);
  n := Inc(a[REAL_TO_INT(r) + 1]);
  n := Two(i := REAL_TO_INT(r), o => x);
  n := REAL_TO_INT(r) + Inc(a[2]);
  Two(o => a[REAL_TO_INT(r)]);
  SPLIT_DATE(IN := D#2024-03-05, YEAR => a[REAL_TO_INT(r)], MONTH => a[1]);
  fs[REAL_TO_INT(r)](d := 1, c := x);
  f(d := 1, c := a[REAL_TO_INT(r)]);
  f(EN := TRUE, d := 1, c := a[REAL_TO_INT(r)], ENO => bs[1]);
  f(d := 1, c := x, q => a[REAL_TO_INT(r)]);
  f(d := 1, c := x, s => ss[REAL_TO_INT(r)]);
  f(d := 1, c := x, ENO => bs[REAL_TO_INT(r)]);
  g(v := aa[REAL_TO_INT(r)]);
  u(f := fs[REAL_TO_INT(r)]);
  tm(IN := TRUE, PT := T#0s, Q => bs[REAL_TO_INT(r)]);
  f(d := 1, c := x, q => a[REAL_TO_INT(r2)]);
  f(d := 1, c := x);
  row := aa[REAL_TO_INT(r)];
  fs[REAL_TO_INT(r)].d := 9;
  rf := REF(a[REAL_TO_INT(r)]);
  q0 := INT_TO_SINT(a[0]);
  q1 := INT_TO_SINT(a[1]);
  q2 := INT_TO_SINT(a[2]);
  q3 := INT_TO_SINT(n);
  q4 := INT_TO_SINT(calls);
  q5 := INT_TO_SINT(f.q);
  q6 := INT_TO_SINT(x);
  q7 := INT_TO_SINT(fs[0].q);
  q8 := INT_TO_SINT(g.n + u.n);
  q9 := INT_TO_SINT(a[3]);
  b0 := bs[0];
  b1 := bs[1];
  b2 := ss[0] = '';
  b3 := tm.Q;
  b4 := rf = NULL;
  q11 := INT_TO_SINT(row[0]);
  q12 := INT_TO_SINT(fs[0].d);
END_PROGRAM

CONFIGURATION c
  VAR_GLOBAL calls : INT; END_VAR
  RESOURCE r ON x
    TASK t(INTERVAL := T#10ms, PRIORITY := 1);
    PROGRAM p WITH t : main;
  END_RESOURCE
END_CONFIGURATION

(* ---- varconfig.st ---- *)
(* AT %I*, %Q*, %M* and VAR_CONFIG (Ed.3 6.5.5.4, 6.4.4.8, 6.8.2): each
   instance's variables where VAR_CONFIG puts them, and initial values
   given per instance, which prevail over the type's. Worked by hand,
   %IW0 2 and %IW2 1 throughout:

   init (cold): hw.out1 and hw2.out1 start at 200 (Q2, Q4: c8 00); lamp
   VAR_CONFIG's 9 (Q1 09) - a `*` address's initial value is given
   there, not where it is declared (Ed.3 Loc_Partly_Var); kept, RETAIN,
   VAR_CONFIG's 60 (M1 3c); t2.out 100 by VAR_CONFIG (Q11 64). Nothing else at a `*`
   address has an initial value: coils, count, arr, t1.out stay 0, and
   an input is the platform's. VAR_CONFIG sets fan.n 10, fan.top 12,
   hw.gain 9.

   tick 0: pump n 1 + 2 = 3, coil 3 > 3 FALSE; fan n 10 + 1 = 11, 11 >
   12 FALSE; st.inner (top 100) n 3, FALSE, st.count 1 (M0); h.v n 1 +
   1 = 2, FALSE: Q0 00. hw.out1 201 (c9 00); hw2 := hw copies the
   values from hw's addresses to hw2's: Q4 c9 00, gain 9. lamp 10, then
   Twice through an in-out: 20 (Q1 14). r := REF(arr[1]), r^ := 300
   (Q8 2c 01); arr[0] := hw2.gain, 9 (Q6 09 00). kept 61 (M1 3d). t1.out
   1, t2.out 101 (Q10 01, Q11 65).
   tick 1: pump n 5 > 3: coil TRUE (Q0 01); fan 12 > 12 FALSE; count 2;
   hw.out1 202 (ca 00), hw2 too; lamp 21, 42 (2a); kept 62; t1 2, t2
   102.
   warm, before tick 2: what is not RETAIN starts again - n 1, top 3,
   out1 200, gain 3 - then VAR_CONFIG's values but kept's, which
   the start keeps (62): fan.n 10, fan.top 12, hw.gain 9, lamp 9,
   t2.out 100. The coils, count, arr and t1.out have no initial value:
   the image keeps them.
   tick 2: pump n 3: coil FALSE (Q0 00); count 3; out1 201; lamp 10,
   20; kept 63 (3f); t1 3, t2 101 (65).
   reference-skip: the reference compiler parses VAR_CONFIG and
   generates nothing for it. *)
TYPE
  HWT : STRUCT
    in1 AT %I* : BOOL;
    out1 AT %Q* : UINT := 200;
    gain : INT := 3;
  END_STRUCT;
  Holder : STRUCT v : valve; END_STRUCT;
END_TYPE
FUNCTION_BLOCK valve
  VAR_INPUT top : INT := 3; END_VAR
  VAR coil AT %Q* : BOOL; level AT %I* : INT; END_VAR
  VAR n : INT := 1; END_VAR
  n := n + level;
  coil := n > top;
END_FUNCTION_BLOCK
FUNCTION_BLOCK station
  VAR inner : valve; END_VAR
  VAR count AT %M* : USINT; END_VAR
  inner(top := 100);
  count := count + 1;
END_FUNCTION_BLOCK
FUNCTION Twice : USINT
  VAR_IN_OUT x : USINT; END_VAR
  x := x * 2;
  Twice := x;
END_FUNCTION
PROGRAM line
  VAR pump, fan : valve; st : station; h : Holder; hw, hw2 : HWT; END_VAR
  VAR lamp AT %Q* : USINT; arr AT %Q* : ARRAY [0..1] OF INT; END_VAR
  VAR RETAIN kept AT %M* : USINT; END_VAR
  VAR r : REF_TO INT; k : USINT; END_VAR
  pump();
  fan();
  st();
  h.v();
  hw.out1 := hw.out1 + 1;
  hw2 := hw;
  lamp := lamp + 1;
  k := Twice(lamp);
  r := REF(arr[1]);
  r^ := 300;
  arr[0] := hw2.gain;
  kept := kept + 1;
END_PROGRAM
PROGRAM tiny
  VAR out AT %Q* : USINT; END_VAR
  out := out + 1;
END_PROGRAM
CONFIGURATION plant
  RESOURCE cpu ON PLC
    TASK fast (INTERVAL := T#10ms, PRIORITY := 1);
    PROGRAM main WITH fast : line;
    PROGRAM t1 WITH fast : tiny;
    PROGRAM t2 WITH fast : tiny;
  END_RESOURCE
  VAR_CONFIG
    cpu.main.pump.coil AT %QX0.0 : BOOL;
    cpu.main.pump.level AT %IW0 : INT;
    cpu.main.fan.coil AT %QX0.1 : BOOL;
    cpu.main.fan.level AT %IW2 : INT;
    cpu.main.fan.n : INT := 10;
    cpu.main.fan.top : INT := 12;
    cpu.main.st.inner.coil AT %QX0.2 : BOOL;
    cpu.main.st.inner.level AT %IW0 : INT;
    cpu.main.st.count AT %MB0 : USINT;
    cpu.main.h.v.coil AT %QX0.3 : BOOL;
    cpu.main.h.v.level AT %IW2 : INT;
    cpu.main.hw.in1 AT %IX4.0 : BOOL;
    cpu.main.hw.out1 AT %QW2 : UINT;
    cpu.main.hw.gain : INT := 9;
    cpu.main.hw2.in1 AT %IX4.1 : BOOL;
    cpu.main.hw2.out1 AT %QW4 : UINT;
    cpu.main.lamp AT %QB1 : USINT := 9;
    cpu.main.arr AT %QW6 : ARRAY [0..1] OF INT;
    cpu.main.kept AT %MB1 : USINT := 60;
    cpu.t1.out AT %QB10 : USINT;
    cpu.t2.out AT %QB11 : USINT := 100;
  END_VAR
END_CONFIGURATION

(* ---- widen.st ---- *)
(* Implicit conversions (Ed.3 6.6.1.6, Figure 11): they widen and keep
   the value - in an assignment, to a block's input and from its output
   (=>), to a function's input, and between the operands of an operator,
   a comparison and MAX; an operation done in its operands' type and
   widened after (Example 3), so INT * INT overflows as an INT even into
   a DINT: at tick 1 30000 * 2 is -5536, flagged.
   Worked by hand: tick 0, vin -3, uin 40000, bin 16#FF, sbin -1: 39997,
   -1, 16#01FF, -1.5, -6, 40001, 200, -4, TRUE, -1. Tick 1, vin 30000,
   uin 2, bin 16#80, sbin 127: 30002, 127, 16#0180, 15000.0, -5536
   (flag), 3, 200, 30127, FALSE, 30000.
   reference-skip: the reference compiler has no implicit conversions
   (Ed.2). *)
FUNCTION_BLOCK pass
VAR_INPUT x : DINT; END_VAR
VAR_OUTPUT y : DINT; o : USINT; END_VAR
y := x + 1;
o := 200;
END_FUNCTION_BLOCK

FUNCTION addl : LINT
VAR_INPUT a : LINT; b : LREAL; END_VAR
addl := a + LREAL_TO_LINT(b);
END_FUNCTION

PROGRAM main
VAR
  vin AT %IW0 : INT;
  uin AT %IW2 : UINT;
  bin AT %IB4 : BYTE;
  sbin AT %IB5 : SINT;
  qd AT %QD0 : DINT;
  ql AT %QL4 : LINT;
  qw AT %QW12 : WORD;
  qr AT %QD14 : REAL;
  qx AT %QD18 : DINT;
  qy AT %QD22 : DINT;
  qo AT %QW26 : INT;
  qf AT %QL28 : LINT;
  qb AT %QX36.0 : BOOL;
  qm AT %QD38 : DINT;
END_VAR
VAR
  d : DINT;
  f : pass;
END_VAR
d := vin;
qd := d + uin;
ql := sbin;
qw := bin OR WORD#16#0100;
qr := vin / REAL#2.0;
qx := vin * 2;
f(x := uin, y => qy, o => qo);
qf := addl(sbin, vin);
qb := d < uin;
qm := MAX(sbin, d);
END_PROGRAM

CONFIGURATION Plant
  RESOURCE r ON PLC
    TASK fast(INTERVAL := T#10ms, PRIORITY := 1);
    PROGRAM p WITH fast : main;
  END_RESOURCE
END_CONFIGURATION

(* ---- wstrings.st ---- *)
(* WSTRING and WCHAR (Ed.3 6.4.2, Tables 6, 25, 27; docs/dependencies.md):
   a WSTRING's characters are UTF-16 units, a character above U+FFFF two
   (a surrogate pair, which LEN counts as two); literals in double quotes
   with $hhhh, ${...}, WCHAR#16#..., and an untyped "X" where a WCHAR is
   wanted (Table 6, 2b); an initial value, in an array and a structure, a
   function block's input and output; CONCAT, LEFT, INSERT, FIND, LEN,
   comparison, s[i] read and written; WORD_TO_WCHAR and WCHAR_TO_WORD
   (binary transfer, Table 25); WSTRING_TO_WCHAR (Table 27 row 2, though
   Figure 11 has none: decided, florin); WSTRING_TO_STRING and
   WCHAR_TO_CHAR, a character a STRING cannot hold skipped, flagged
   CONVERSION; INT_TO_WSTRING and WSTRING_TO_INT.
   Worked by hand, the input wc:
   tick 0, 'q' (16#0071): ws "a$263Aq", t "a$263Aqz": qlen 16#24 (LEN(t) 4,
   LEN(emoji) 2), qfind 4, qc 16#263A, qcmp TRUE, qeq TRUE, qn 75, qs '<q>',
   qch 'q', qw 16#0061, qk 4, qr 'q' (r.w "hqi"), qx 'q' (k.last[3]).
   Tick 1, 16#00E9 (e acute, in Latin-1): the same with 16#E9; qs '<'
   16#E9 '>'.
   Tick 2, 16#4E2D (a CJK character): qs '<>', qch '$00', qr and qx
   16#4E2D; flagged CONVERSION at line 75 (WSTRING_TO_STRING), the first
   flag, which stays until the platform clears it (docs/c-output.md §5).
   Tick 3, 16#0030 ('0'): WSTRING_TO_WCHAR of an empty WSTRING, "$0000"
   into qx (flagged too, behind the flag of tick 2: the book's checked
   table shows that flag, docs/behaviour/strings.md).
   reference-skip: WCHAR and s[i] are Ed.3's; the reference compiler
   (Ed.2) has neither. *)
TYPE rec : STRUCT w : WSTRING[4] := "hi"; c : WCHAR := "z"; END_STRUCT; END_TYPE

FUNCTION_BLOCK keep
VAR_INPUT s : WSTRING[8]; END_VAR
VAR_OUTPUT last : WSTRING[8] := "?"; n : INT; END_VAR
last := s;
n := LEN(s);
END_FUNCTION_BLOCK

PROGRAM main
VAR
  win AT %IW0 : WORD;
  qlen AT %QB0 : USINT;
  qfind AT %QB1 : USINT;
  qc AT %QW2 : WCHAR;
  qcmp AT %QX4.0 : BOOL;
  qeq AT %QX4.1 : BOOL;
  qn AT %QB5 : USINT;
  qs AT %QB6 : STRING[6];
  qch AT %QB13 : CHAR;
  qw AT %QW14 : WORD;
  qk AT %QB16 : USINT;
  qr AT %QW17 : WCHAR;
  qx AT %QW19 : WCHAR;
END_VAR
VAR
  ws : WSTRING[6] := "a$263Ab";
  wc : WCHAR;
  emoji : WSTRING := "${1F600}";
  arr : ARRAY[0..1] OF WSTRING[3] := ["xy", "z"];
  r : rec;
  k : keep;
  t : WSTRING[6];
  e : WSTRING[2] := "";
END_VAR
wc := WORD_TO_WCHAR(win);
ws[3] := wc;
t := CONCAT(ws, arr[1]);
qlen := INT_TO_USINT(LEN(t)) + INT_TO_USINT(LEN(emoji)) * 16;
qfind := INT_TO_USINT(FIND(t, "z"));
qc := t[2];
qcmp := t > "a";
qeq := LEFT(t, 1) = "a" AND r.c = "z";
qn := INT_TO_USINT(WSTRING_TO_INT(CONCAT(INT_TO_WSTRING(7), "5")));
k(s := t);
qk := INT_TO_USINT(k.n);
r.w := "hi";
r.w := INSERT(r.w, wc, 1);
qr := r.w[2];
qs := WSTRING_TO_STRING(CONCAT("<", wc, ">"));
qch := WCHAR_TO_CHAR(wc);
qw := WCHAR_TO_WORD(WSTRING_TO_WCHAR(t));
IF wc = "0" THEN
  qx := WSTRING_TO_WCHAR(e);
ELSE
  qx := k.last[3];
END_IF;
END_PROGRAM

CONFIGURATION Plant
  RESOURCE r ON PLC
    TASK fast(INTERVAL := T#10ms, PRIORITY := 1);
    PROGRAM p WITH fast : main;
  END_RESOURCE
END_CONFIGURATION

(* ---- arith.st ---- *)
(* Integer arithmetic of every width, in range: + - * / MOD, negation,
   ABS, MIN, MAX, LIMIT, and division and MOD of negative numbers. *)
PROGRAM main
VAR
  a AT %IW0 : INT;
  b AT %IW2 : INT;
  r_add AT %MW0 : INT;
  r_sub AT %MW2 : INT;
  r_mul AT %MD4 : DINT;
  r_div AT %MW8 : INT;
  r_mod AT %MW10 : INT;
  r_neg AT %MW12 : INT;
  r_abs AT %MW14 : INT;
  r_min AT %MW16 : INT;
  r_max AT %MW18 : INT;
  r_lim AT %MW20 : INT;
  s AT %MB22 : SINT;
  us AT %MB23 : USINT;
  ui AT %MW24 : UINT;
  ud AT %MD26 : UDINT;
  l AT %ML30 : LINT;
  ul AT %ML38 : ULINT;
END_VAR
r_add := a + b;
r_sub := a - b;
r_mul := INT_TO_DINT(a) * INT_TO_DINT(b);
IF b <> 0 THEN
  r_div := a / b;
  r_mod := a MOD b;
END_IF;
r_neg := -a;
r_abs := ABS(a);
r_min := MIN(a, b, 7);
r_max := MAX(a, b, -7);
r_lim := LIMIT(-100, a * 3, 100);
s := INT_TO_SINT(a) - SINT#3;
us := USINT#200 + USINT#5;
ui := UINT#60000 / UINT#7;
ud := UDINT#4000000000 - UDINT#1;
l := INT_TO_LINT(a) * LINT#1000000000000;
ul := ULINT#18000000000000000000 + INT_TO_ULINT(ABS(b));
END_PROGRAM

CONFIGURATION plant
  RESOURCE r ON PLC
    TASK fast(INTERVAL := T#10ms, PRIORITY := 0);
    PROGRAM p WITH fast : main;
  END_RESOURCE
END_CONFIGURATION

(* ---- autoaddr.st ---- *)
(* TwinCAT's automatic addressing (auto-addresses): a `*` address no
   VAR_CONFIG entry gives - a global's own, a global's `*` components,
   a program instance's - placed by iecf in its area after the last
   byte any stated address reaches, in the order of the paths, each its
   own type's width, a BOOL a whole byte.
   Stated: x AT %MW10 (M up to 12), VAR_CONFIG RS.P.D.Q AT %QW20 (Q up
   to 22). Placed, by path: I: DEV.A 0, RS.P.D.A 2. Q: DEV.Q 22, FLAG
   24. M: ARR 12 (4 bytes), DEV.M 16, G 18, RS.P.D.M 20, RS.P.P 22.
   Worked by hand, each tick: g + 1, dev.m + 2, p + 3, flag TRUE,
   dev.q := g * 10, arr[1] + 7, d.q := 5, d.m + 1, x + 100.
   Tick 1: M x 100, arr 0 7, dev.m 2, g 1, d.m 1, p 3; Q d.q 5,
   dev.q 10, flag 1. Tick 2: x 200, arr 0 14, dev.m 4, g 2, d.m 2,
   p 6; d.q 5, dev.q 20, flag 1.
   reference-skip: not IEC 61131-3. *)
TYPE Io : STRUCT
  a AT %I* : INT;
  q AT %Q* : INT;
  m AT %M* : INT;
END_STRUCT;
END_TYPE

PROGRAM main
  VAR p AT %M* : INT; END_VAR
  VAR d : Io; END_VAR
  VAR x AT %MW10 : INT; END_VAR
  VAR_EXTERNAL g : INT; flag : BOOL; dev : Io; arr : ARRAY[0..1] OF INT; END_VAR
  g := g + 1;
  dev.m := dev.m + 2;
  p := p + 3;
  flag := TRUE;
  dev.q := g * 10;
  arr[1] := arr[1] + 7;
  d.q := 5;
  d.m := d.m + 1;
  x := x + 100;
END_PROGRAM

CONFIGURATION cf
  VAR_GLOBAL
    g AT %M* : INT;
    flag AT %Q* : BOOL;
    arr AT %M* : ARRAY[0..1] OF INT;
  END_VAR
  VAR_GLOBAL
    dev : Io;
  END_VAR
  RESOURCE rs ON x
    TASK tk(INTERVAL := T#10ms, PRIORITY := 1);
    PROGRAM p WITH tk : main;
  END_RESOURCE
  VAR_CONFIG
    rs.p.d.q AT %QW20 : INT;
  END_VAR
END_CONFIGURATION

(* ---- bcd.st ---- *)
(* BCD conversions (Ed.3 6.6.2.5.2, Table 22 3a-4b, footnote d), by the
   names the reference compiler has too. Each nibble a decimal digit, the
   lowest the units. Inputs w (%IW0) and u (%IW2), so nothing is folded.
   Worked by hand:
   tick 0, w 16#0099, u 1234: a := WORD_BCD_TO_UINT(w) 99 (63 00);
     b := UINT_TO_BCD_WORD(u) 16#1234 (34 12); c, of w's low byte, 99
     (63); d := USINT_TO_BCD_BYTE(34) 16#34; e, of 16#12340099,
     12340099 (83 4b bc 00); f := ULINT_TO_BCD_LWORD(u * 10^11)
     16#0123400000000000; g := BCD_TO_UINT(w), the overloaded form, 99;
     h := WORD_BCD_TO_USINT(w) 99; k, f back, 123400000000000.
   tick 1, w 16#12A4, u 10000: w is not BCD (a nibble A), so a, c, e, g
     and h are 0, as the reference compiler gives (its ENO FALSE); iecf
     also flags it, "flag 4 MAIN 37" at a, the first. u has five digits,
     more than a WORD's four: b is every nibble F, 16#FFFF (ff ff),
     where the reference compiler keeps the low digits, 16#0000: iecf's
     choice, so its bytes are bcd.iecf.trace's (docs/dependencies.md). f is
     16#1000000000000000, k 10^15.
   tick 2, w 16#9999, u 99: a 9999 (0f 27), b 16#0099, c 99, d 16#99,
     e 12349999, f 16#0009900000000000, g 9999; h 9999 is beyond USINT,
     which keeps its low bits as any conversion does: 15 (0f). *)
PROGRAM main
VAR
  w AT %IW0 : WORD;
  u AT %IW2 : UINT;
END_VAR
VAR
  a AT %MW0 : UINT;
  b AT %MW2 : WORD;
  c AT %MB4 : USINT;
  d AT %MB5 : BYTE;
  e AT %MD6 : UDINT;
  f AT %ML10 : LWORD;
  g AT %MW18 : UINT;
  h AT %MB20 : USINT;
  k AT %ML24 : ULINT;
END_VAR
a := WORD_BCD_TO_UINT(w);
b := UINT_TO_BCD_WORD(u);
c := BYTE_BCD_TO_USINT(WORD_TO_BYTE(w));
d := USINT_TO_BCD_BYTE(UINT_TO_USINT(u MOD 100));
e := DWORD_BCD_TO_UDINT(WORD_TO_DWORD(w) OR 16#12340000);
f := ULINT_TO_BCD_LWORD(UINT_TO_ULINT(u) * 100000000000);
g := BCD_TO_UINT(w);
h := WORD_BCD_TO_USINT(w);
k := LWORD_BCD_TO_ULINT(f);
END_PROGRAM

CONFIGURATION Plant
  RESOURCE R ON PLC
    TASK fast(INTERVAL := T#10ms, PRIORITY := 1);
    PROGRAM P WITH fast : main;
  END_RESOURCE
END_CONFIGURATION
